(* IEC 61131-3 sources: JingjiangMoonbox/Application/Application/任务列表/Main_Task/IO列表, 15 files *)

(* ---- StEvtReq.st ---- *)
(*@CES
Name=StEvtReq
Type=Gvl
TypeGuid=2db5746d-d284-4425-9f7f-2663a34b0ebc
Guid=8252279d-9d67-4d9b-8f5c-5fb7a358024a
HasDeclaration=True
HasImplementation=False
*)
{DECLARATION}
{attribute 'pack_mode' := '1'}
TYPE StEvtReq :
STRUCT
	xEvt_Estop						: BOOL; (* 急停 *)
	xEvt_Stop						: BOOL; (* 停机 *)
	xEvt_Tension					: BOOL; (* 张力投入 *)
	xEvt_ManuSpdUp					: BOOL; (* 手动加速 *)
	xEvt_ManuSpdDn					: BOOL; (* 手动减速 *)
	xEvt_Ink						: BOOL; (* 空转 *)
	xEvt_Prestart					: BOOL; (* (预)启动 *)
	xEvt_PressAll					: BOOL; (* 全体合压 *)
	xEvt_UnpressAll					: BOOL; (* 全体离压 *)
	xEvt_Print						: BOOL; (* 印刷|联动 *)
	xEvt_AlarmBell					: BOOL; (* 报警 *)
	xEvt_AllInchRun					: BOOL; (* 整机单动 *)
	xEvt_AllExhBlower				: BOOL; (* 整机排风 *)
	xEvt_AllCoolBlower				: BOOL; (* 整机冷风 *)
	xEvt_AllHotBlower				: BOOL; (* 整机热风 *)
	xEvt_AllHeating					: BOOL; (* 整机加热 *)
	xEvt_TapPosition_Printing		: BOOL; (* 2018.7.16.151840/印刷档位 *)
	xEvt_TapPosition_Breaking		: BOOL; (* 2018.7.16.151514/断料档位 *)
	xEvt_TapPosition_UniformInk		: BOOL; (* 2018.7.16.151507/匀墨档位 *)
	xEvt_FastStop					: BOOL;	(* 2022.4.6.110418 快停*)

	xReqEstop						: BOOL; (* 急停 *)
	xReqStop						: BOOL; (* 停机 *)
	xReqTension						: BOOL; (* 张力投入 *)
	xReqManuSpdUp					: BOOL; (* 手动加速 *)
	xReqManuSpdDn					: BOOL; (* 手动减速 *)
	xReqInk							: BOOL; (* 空转 *)
	xReqPrestart					: BOOL; (* (预)启动 *)
	xReqPressAll					: BOOL; (* 全体合压 *)
	xReqUnpressAll					: BOOL; (* 全体离压 *)
	xReqPrint						: BOOL; (* 印刷|联动 *)
	xReqAlarmBell					: BOOL; (* 报警 *)
	xReqAllInchRun					: BOOL; (* 整机单运行 *)
	xReqAllExhBlower				: BOOL; (* 整机排风 *)
	xReqAllCoolBlower				: BOOL; (* 整机冷风 *)
	xReqAllHotBlower				: BOOL; (* 整机热风 *)
	xReqAllHeating					: BOOL; (* 整机加热 *)
	xReqFastStop					: BOOL;	(* 2022.4.6.110418 快停*)
END_STRUCT
END_TYPE

{IMPLEMENTATION}

(* ---- StIOMap_Axis_Extra_FE.st ---- *)
(*@CES
Name=StIOMap_Axis_Extra_FE
Type=Gvl
TypeGuid=2db5746d-d284-4425-9f7f-2663a34b0ebc
Guid=0a3c1562-979e-4c29-a397-fc51d923e0fc
HasDeclaration=True
HasImplementation=False
*)
{DECLARATION}
{attribute 'pack_mode' := '1'}
TYPE StIOMap_Axis_Extra_FE :
STRUCT
	i_xPreHeating							: BOOL; (* 预加热 *)
	i_xPreHeating_Err						: BOOL; (* 预加热报警\温控信号 *)
	i_xPreHotBlower							: BOOL; (* 预热风 *)
	i_xPreHotBlower_Err						: BOOL; (* 预热风报警 *)
	i_xCoolBlower							: BOOL; (* 冷风开关 *)
	i_xCoolBlower_Button					: BOOL; (* 冷风按钮 *)
	i_xCoolBlower_Err						: BOOL; (* 冷风报警 *)
	i_xHotBlower							: BOOL; (* 热风开关 *)
	i_xHotBlower_Button						: BOOL; (* 热风按钮 *)
	i_xHotBlower_Err						: BOOL; (* 热风报警 *)
	i_xHotBlower_Opened_Act					: BOOL; (* 热风实际被打开了|2022.5.11.192858|没有反馈时候需要写true*)
	i_xHotBlower_CHNL2						: BOOL; (* 第2路热风开关 *)
	i_xHotBlower_Button_CHNL2				: BOOL; (* 第2路热风按钮 *)
	i_xHotBlower_Err_CHNL2					: BOOL; (* 第2路热风报警 *)
	i_xHotBlower_Opened_Act_CHNL2			: BOOL; (* 热风2实际被打开了|2022.5.11.192858|没有反馈时候需要写true*)
	i_xTemReachToTarget						: BOOL; (* 到达目标温度 *)
	i_xSteamHeating							: BOOL; (* 蒸汽加热开关 *)
	i_xSteamHeating_Err						: BOOL; (* 蒸汽加热报警 *)
	i_xHeating_I							: BOOL; (* 电加热I档 *)
	i_xHeating_II							: BOOL; (* 电加热II档 *)
	i_xHeating_III							: BOOL; (* 电加热III档 *)
	i_xHeating_Button						: BOOL; (* 加热按钮 *)
	i_xHeating_I_CHNL2						: BOOL; (* 第2路电加热I档 *)
	i_xHeating_II_CHNL2						: BOOL; (* 第2路电加热II档 *)
	i_xHeating_III_CHNL2					: BOOL; (* 第2路电加热III档 *)
	i_xHeating_Button_CHNL2					: BOOL; (* 第2路加热按钮 *)
	i_xAllExhBlower_Up						: BOOL; (* 全上排风 *)
	i_xAllExhBlower_Err_Up					: BOOL; (* 上排风报警 *)
	i_xAllExhBlower_Dn						: BOOL; (* 全下排风 *)
	i_xAllExhBlower_Err_Dn					: BOOL; (* 下排风报警 *)
	i_xAllCoolBlower						: BOOL; (* 全冷风 *)
	i_xAllHotBlower							: BOOL; (* 全热风 *)
	i_xAllHeating							: BOOL; (* 全加热 *)
	i_xAirInletMotorMin_Limit				: BOOL; (* 进风口风门电机最小开度限位 *)
	i_xAirInletMotorMax_Limit				: BOOL; (* 进风口风门电机最大开度限位 *)
	i_xOvensAirOutMotorMin_Limit			: BOOL; (* 烘箱出风口风门电机最小开度限位 *)
	i_xOvensAirOutMotorMax_Limit			: BOOL; (* 烘箱出风口风门电机最大开度限位 *)
	i_xAirExhaustMotorMin_Limit				: BOOL; (* 排风口风门电机最小开度限位 *)
	i_xAirExhaustMotorMax_Limit				: BOOL; (* 排风口风门电机最大开度限位 *)
	i_xAirReturnMotorMin_Limit				: BOOL; (* 回风口风门电机最小开度限位 *)
	i_xAirReturnMotorMax_Limit				: BOOL; (* 回风口风门电机最大开度限位 *)
	i_xScraperInveterError					: BOOL; (* 刮刀变频器报警 *)
	i_xScraperOn							: BOOL; (* 刮刀开关 *)
	i_xInkRollerInveterError				: BOOL; (* 递墨辊变频器报警 |2022.3.26.094940*)
	i_xInkRoller_CW							: BOOL; (* 递墨辊正转开 *)
	i_xInkRoller_CCW						: BOOL; (* 递墨辊反转开 *)
	i_xInkRoller_Up							: BOOL; (* 递墨辊上 *)
	i_xInkRoller_Dn							: BOOL; (* 递墨辊下 *)
	i_xTurnoverFilmAgency					: BOOL; (* 翻料架开关 *)
	i_wAI_AirInletMotor						: WORD; (* 进风口反馈|模拟量控制风门LEL *)
	i_wAI_OvensAirOutMotor					: WORD; (* 烘箱出风口反馈|模拟量控制风门LEL *)
	i_wAI_AirExhaustMotor					: WORD; (* 排风口反馈|模拟量控制风门LEL *)
	i_wAI_AirReturnMotor					: WORD; (* 回风反馈|模拟量控制风门LEL *)
	i_wInputLel								: WORD; (* LEL浓度反馈 *)
	i_wInAllAir								: WORD; (* 总进风反馈输入 *)
	i_wInFreshAir							: WORD; (* 新风反馈输入 *)
	i_wInExhaustAir							: WORD; (* 排风反馈输入 *)
	i_wInReturnAir							: WORD; (* 二次回风反馈输入 *)
	i_xTaper_Incr							: BOOL; (* 增加锥度+|针对牵引 *)
	i_xTaper_Decr							: BOOL; (* 减小锥度-|针对牵引 *)
	i_wAI_CoatingSensor						: WORD; (* 涂布传感器模拟量 *)
	i_byAIType_CoatingSensor				: BYTE; (* 涂布传感器类型 *)
	i_xAirExhaustSwitch						: BOOL; (* 色组排风输入开关 *)
	i_xAirExhaustButton						: BOOL; (* 色组排风输入按钮 *)
	i_xPushIn_PrnRoller						: BOOL; (* 顶版-进 *)
	i_xPullOut_PrnRoller					: BOOL; (* 顶版-退 *)
	i_xRsvd_DI0								: BOOL; (* 数字量输入保留0 *)
	i_xRsvd_DI1								: BOOL; (* 数字量输入保留1 *)
	i_xRsvd_DI2								: BOOL; (* 数字量输入保留2 *)
	i_xRsvd_DI3								: BOOL; (* 数字量输入保留3 *)
	i_xRsvd_DI4								: BOOL; (* 数字量输入保留4 *)
	i_xRsvd_DI5								: BOOL; (* 数字量输入保留5 *)
	i_xRsvd_DI6								: BOOL; (* 数字量输入保留6 *)
	i_xRsvd_DI7								: BOOL; (* 数字量输入保留7 *)
	i_xRsvd_DI8								: BOOL; (* 数字量输入保留8 *)
	i_xRsvd_DI9								: BOOL; (* 数字量输入保留9 *)
	i_xRsvd_DI10							: BOOL; (* 数字量输入保留10 *)
	i_xRsvd_DI11							: BOOL; (* 数字量输入保留11 *)
	i_xRsvd_DI12							: BOOL; (* 数字量输入保留12 *)
	i_xRsvd_DI13							: BOOL; (* 数字量输入保留13 *)
	i_xRsvd_DI14							: BOOL; (* 数字量输入保留14 *)
	i_xRsvd_DI15							: BOOL; (* 数字量输入保留15 *)
	i_wRsvd_AI0								: WORD; (* 模拟量输入保留0 *)
	i_wRsvd_AI1								: WORD; (* 模拟量输入保留1 *)
	i_wRsvd_AI2								: WORD; (* 模拟量输入保留2 *)
	i_wRsvd_AI3								: WORD; (* 模拟量输入保留3 *)
	i_wRsvd_AI4								: WORD; (* 模拟量输入保留4 *)
	i_wRsvd_AI5								: WORD; (* 模拟量输入保留5 *)

	o_xRel_PreHeating						: BOOL; (* 预加热接触器 *)
	o_xLamp_PreHeating						: BOOL; (* 预加热指示灯 *)
	o_xRel_ResetErr_PreHeating				: BOOL; (* 预加热故障复位 *)
	o_wAO_PreHeating						: WORD; (* 预加热模拟量 *)
	o_xRel_PreHeatingRoller_Motor			: BOOL; (* 预热辊使能 *)
	o_xRel_PreHeatingRoller_Motor_Rev		: BOOL; (* 预热辊反转使能 *)
	o_wAO_PreHeatingRoller_Motor			: WORD; (* 预热辊模拟量输出 *)
	o_xRel_PreHotBlower						: BOOL; (* 预热风接触器 *)
	o_xLamp_PreHotBlower					: BOOL; (* 预热风指示灯 *)
	o_xRel_ResetErr_PreHotBlower			: BOOL; (* 预热风故障复位 *)
	o_wAO_PreHotBlower						: WORD; (* 预热风模拟量 *)
	o_xRel_CoolBlower						: BOOL; (* 冷风接触器 *)
	o_xLamp_CoolBlower						: BOOL; (* 冷风指示灯 *)
	o_xRel_HotBlower						: BOOL; (* 热风接触器 *)
	o_xLamp_HotBlower						: BOOL; (* 热风指示灯 *)
	o_xRel_ResetErr_HotBlower				: BOOL; (* 热风故障复位 *)
	o_wAO_HotBlower							: WORD; (* 热风模拟量输出 *)
	o_xRel_HotBlower_CHNL2					: BOOL; (* 第2路热风接触器 *)
	o_xLamp_HotBlower_CHNL2					: BOOL; (* 第2路热风指示灯 *)
	o_xRel_ResetErr_HotBlower_CHNL2			: BOOL; (* 第2路热风故障复位 *)
	o_wAO_HotBlower_CHNL2					: WORD; (* 第2路热风模拟量输出 *)
	o_xRel_SteamHeating						: BOOL; (* 蒸汽输出 *)
	o_xLamp_SteamHeating					: BOOL; (* 蒸汽加热指示灯 *)
	o_xRel_ResetErr_SteamHeating			: BOOL; (* 蒸汽加热复位 *)
	o_wAO_SteamHeating						: WORD; (* 蒸汽加热模拟量输出 *)
	o_xRel_Heating_I						: BOOL; (* 电加热I档 *)
	o_xRel_Heating_II						: BOOL; (* 电加热II档 *)
	o_xRel_Heating_III						: BOOL; (* 电加热III档 *)
	o_xLamp_Heating							: BOOL; (* 电加热指示灯 *)
	o_xRel_Heating_I_CHNL2					: BOOL; (* 第2路电加热I档 *)
	o_xRel_Heating_II_CHNL2					: BOOL; (* 第2路电加热II档 *)
	o_xRel_Heating_III_CHNL2				: BOOL; (* 第2路电加热III档 *)
	o_xLamp_Heating_CHNL2					: BOOL; (* 第2路电加热指示灯 *)
	o_xRel_AllExhBlower_Up					: BOOL; (* 上排风继电器输出 *)
	o_xLamp_AllExhBlower_Up					: BOOL; (* 全上排风指示灯 *)
	o_xRel_ModeStar_AllExhBlower_Up			: BOOL; (* 上排风模式-星形 *)
	o_xRel_ModeTriangle_AllExhBlower_Up		: BOOL; (* 上排风模式-三角 *)
	o_xRel_ResetErr_AllExhBlower_Up			: BOOL; (* 上排风故障复位 *)
	o_wAO_AllExhBlower_Up					: WORD; (* 上排风模拟量输出 *)
	o_xRel_AllExhBlower_Dn					: BOOL; (* 下排风继电器输出 *)
	o_xLamp_AllExhBlower_Dn					: BOOL; (* 全下排风指示灯 *)
	o_xRel_ModeStar_AllExhBlower_Dn			: BOOL; (* 下排风模式-星形 *)
	o_xRel_ModeTriangle_AllExhBlower_Dn		: BOOL; (* 下排风模式-三角 *)
	o_xRel_ResetErr_AllExhBlower_Dn			: BOOL; (* 下排风故障复位 *)
	o_wAO_AllExhBlower_Dn					: WORD; (* 下排风模拟量输出 *)
	o_xLamp_AllCoolBlower					: BOOL; (* 全冷风指示灯 *)
	o_xLamp_AllHotBlower					: BOOL; (* 全热风指示灯 *)
	o_xLamp_AllHeating						: BOOL; (* 全加热指示灯 *)
	o_xAirInletMotor_Increase				: BOOL; (* 进风口风门开度增大 *)
	o_xAirInletMotor_Decrease				: BOOL; (* 进风口风门开度减小 *)
	o_xOvensAirOutMotor_Increase			: BOOL; (* 烘箱出风口风门开度增大 *)
	o_xOvensAirOutMotor_Decrease			: BOOL; (* 烘箱出风口风门开度减小 *)
	o_xAirExhaustMotor_Increase				: BOOL; (* 排风口风门开度增大 *)
	o_xAirExhaustMotor_Decrease				: BOOL; (* 排风口风门开度减小 *)
	o_xAirReturnMotor_Increase				: BOOL; (* 回风风门开度增大 *)
	o_xAirReturnMotor_Decrease				: BOOL; (* 回风风门开度减小 *)
	o_xScraperOn							: BOOL; (* 刮刀输出 *)
(*2022.7.8.093123*)
	o_xScraperRst							: BOOL;(*刮刀故障复位*)
	o_wAO_Scraper							: WORD; (* 刮刀模拟量输出 *)
	o_xInkRollerOn							: BOOL; (* 递墨辊运动信号 *)
	o_xInkRollerRst							: BOOL;(*递墨辊复位2022.7.8.093223*)
	o_xRel_InkRoller_CW						: BOOL; (* 递墨辊正转 *)
	o_xRel_InkRoller_CCW					: BOOL; (* 递墨辊反转 *)
	o_wAO_InkRoller							: WORD; (* 递墨辊模拟量输出 *)
	(*2026.05.25.134825*)
	o_wAO_InkRoller_Dir						:WORD;(*递墨辊模拟量输出@±10V*)
	o_xRel_InkRoller_Up						: BOOL; (* 递墨辊上输出 *)
	o_xRel_InkRoller_Dn						: BOOL; (* 递墨辊下输出 *)
	o_xRel_TurnoverFilmAgency				: BOOL; (* 翻料架输出 *)
	o_xRel_ColdWaterRoller_Motor			: BOOL; (* 水冷辊电机使能 *)
	o_xRel_ColdWaterRoller_Motor_Rev		: BOOL; (* 水冷辊电机反转使能 *)
	o_wAO_ColdWaterRoller_Motor				: WORD; (* 水冷辊电机模拟量输出 *)
	o_xRel_DriveAfterPrint_Motor			: BOOL; (* 印后传动辊电机使能 *)
	o_xRel_DriveAfterPrint_Motor_Rev		: BOOL; (* 印后传动辊电机反转 *)
	o_wAO_DriveAfterPrint_Motor				: WORD; (* 印后传动辊电机模拟量输出 *)
	o_wAO_AirInletMotor						: WORD; (* 进口输出|模拟量控制风门LEL *)
	o_wAO_OvensAirOutMotor					: WORD; (* 烘箱出风口输出|模拟量控制风门LEL *)
	o_wAO_AirExhaustMotor					: WORD; (* 排风口输出|模拟量控制风门LEL *)
	o_wAO_AirReturnMotor					: WORD; (* 回风输出|模拟量控制风门LEL *)
	o_wInAllAir								: WORD; (* 总进风输出 *)
	o_wInFreshAir							: WORD; (* 新风输出 *)
	o_wInExhaustAir							: WORD; (* 排风输出 *)
	o_wInReturnAir							: WORD; (* 二次回风输出 *)
	o_wPreAirHotRollTorque					: WORD; (* 预热辊转矩输出 *)
	o_wCoolWaterRollTorque					: WORD; (* 水冷辊转矩输出 *)
	o_xAirExhaustEn							: BOOL; (* 色组排风输出使能 *)
	o_xRel_PushIn_PrnRoller					: BOOL; (* 顶版-进执行 *)
	o_xRel_PullOut_PrnRoller				: BOOL; (* 顶版-退执行 *)
	o_xRel_ModeStar_HotBlower				: BOOL; (* 热风输出-星形 *)
	o_xRel_ModeTriangle_HotBlower			: BOOL; (* 热风输出-三角 *)
	o_xRel_Oven								: BOOL; (* 色组烘箱输出 *)
	o_xRsvd_DO0								: BOOL; (* 数字量输出保留0 *)
	o_xRsvd_DO1								: BOOL; (* 数字量输出保留1 *)
	o_xRsvd_DO2								: BOOL; (* 数字量输出保留2 *)
	o_xRsvd_DO3								: BOOL; (* 数字量输出保留3 *)
	o_xRsvd_DO4								: BOOL; (* 数字量输出保留4 *)
	o_xRsvd_DO5								: BOOL; (* 数字量输出保留5 *)
	o_xRsvd_DO6								: BOOL; (* 数字量输出保留6 *)
	o_xRsvd_DO7								: BOOL; (* 数字量输出保留7 *)
	o_xRsvd_DO8								: BOOL; (* 数字量输出保留8 *)
	o_xRsvd_DO9								: BOOL; (* 数字量输出保留9 *)
	o_xRsvd_DO10							: BOOL; (* 数字量输出保留10 *)
	o_xRsvd_DO11							: BOOL; (* 数字量输出保留11 *)
	o_xRsvd_DO12							: BOOL; (* 数字量输出保留12 *)
	o_xRsvd_DO13							: BOOL; (* 数字量输出保留13 *)
	o_xRsvd_DO14							: BOOL; (* 数字量输出保留14 *)
	o_xRsvd_DO15							: BOOL; (* 数字量输出保留15 *)
	o_wRsvd_AO0								: WORD; (* 模拟量输出保留0 *)
	o_wRsvd_AO1								: WORD; (* 模拟量输出保留1 *)
	o_wRsvd_AO2								: WORD; (* 模拟量输出保留2 *)
	o_wRsvd_AO3								: WORD; (* 模拟量输出保留3 *)
	o_wRsvd_AO4								: WORD; (* 模拟量输出保留4 *)
	o_wRsvd_AO5								: WORD; (* 模拟量输出保留5 *)
END_STRUCT
END_TYPE

{IMPLEMENTATION}

(* ---- StIOMap_Axis_FE.st ---- *)
(*@CES
Name=StIOMap_Axis_FE
Type=Gvl
TypeGuid=2db5746d-d284-4425-9f7f-2663a34b0ebc
Guid=869f751a-dcb2-42ff-ace2-93e211c33fe9
HasDeclaration=True
HasImplementation=False
*)
{DECLARATION}
{attribute 'pack_mode' := '1'}
TYPE StIOMap_Axis_FE :
STRUCT
	(*IO输入*)
	i_xLinkage								: BOOL; (* 联动 *)
	i_xInch									: BOOL; (* 单运行 *)
	i_xEstop								: BOOL; (* 急停输入 *)
	i_xAlarmBell							: BOOL; (* 警报 *)
	i_xBigAdj								: BOOL; (* 粗调 *)
	i_xLittleAdj							: BOOL; (* 细调 *)
	i_xPressMode_Auto						: BOOL; (* 自动合压 *)
	i_xPressMode_Manu						: BOOL; (* 手动合压 *)
	i_xPress								: BOOL; (* 合压输入 *)
	i_xUnPress								: BOOL; (* 离压输入 *)
	i_xUnPress_Inching						: BOOL; (* 点动离压 *)
	i_xMove_Up								: BOOL; (* 上调 *)
	i_xMove_Down							: BOOL; (* 下调 *)
	i_xMove_Left							: BOOL; (* 左调 *)
	i_xMove_Right							: BOOL; (* 右调 *)
	i_xPosLimit_Left						: BOOL; (* 左限位 *)
	i_xPosLimit_Right						: BOOL; (* 右限位 *)
	i_xHorzMotor_FastSpd					: BOOL; (* 横向电机快 *)
	i_xSleeve_Prn							: BOOL; (* 版辊套筒*)
	i_xSleeve_Net							: BOOL; (* 网辊套筒*)
	i_xPlate_Push_Prn						: BOOL; (* 版辊推出*)
	i_xPlate_Push_Net						: BOOL; (* 网辊推出*)
	i_xAcc									: BOOL; (* 加速 *)
	i_xDec									: BOOL; (* 减速 *)
	i_xInch_Net								: BOOL; (* 网辊单运行-匀墨 *)
		(*2024.09.28.094834//增加秦华IO*)
	i_xJogPaper									: BOOL; (* 走纸点动 *)
	i_xEn_Prn									: BOOL; (* 版辊使能开关 *)

	i_xPrnBigAdj								: BOOL; (* 印刷辊粗调 *)
	i_xPrnLittleAdj								: BOOL; (* 印刷辊细调 *)
	i_xNetBigAdj								: BOOL; (* 网辊粗调 *)
	i_xNetLittleAdj								: BOOL; (* 网辊细调 *)
	i_xStrBigAdj								: BOOL; (* 张带辊粗调 *)
	i_xStrLittleAdj								: BOOL; (* 张带辊细调 *)

	i_xJogUp_Prn_M							: BOOL; (* 印刷辊点动上升 *)
	i_xJogDown_Prn_M						: BOOL; (* 印刷辊点动下降 *)
	i_xJogUp_Prn_G							: BOOL; (* 印刷辊点进上升  传动侧信号*)
	i_xJogDown_Prn_G						: BOOL; (* 印刷辊点动下降  传动侧信号*)
	i_xAllUp_Prn							: BOOL; (* 印刷辊整体上升 *)
	i_xAllDown_Prn							: BOOL; (* 印刷辊整体下降 *)
	i_xJogUp_Str_M							: BOOL; (* 张带辊点动上升 *)
	i_xJogDown_Str_M						: BOOL; (* 张带辊点动下降 *)
	i_xJogUp_Str_G							: BOOL; (* 张带辊点动上升  传动侧信号*)
	i_xJogDown_Str_G						: BOOL; (* 张带辊点动下降  传动侧信号*)
	i_xAllUp_Str							: BOOL; (* 张带辊整体上升 *)
	i_xAllDown_Str							: BOOL; (* 张带辊整体下降 *)
	i_xJogUp_Net_M							: BOOL; (* 网版辊点动前进 *)
	i_xJogDown_Net_M						: BOOL; (* 网版辊点动后退 *)
	i_xJogUp_Net_G							: BOOL; (* 网版辊点动前进 另传动侧信号*)
	i_xJogDown_Net_G						: BOOL; (* 网版辊点动后退  另传动侧信号*)
	i_xAllUp_Net							: BOOL; (* 网版辊整体前进 *)
	i_xAllDown_Net							: BOOL; (* 网版辊整体后退 *)

	i_xSuctionMotor							: BOOL; (* 吸风电机开关*)
	i_xNetMotor								: BOOL;(* 网辊电机开关*)
	i_xNetLock								: BOOL;(* 网辊锁紧开关*)
	i_xStop                             	: BOOL;(* 停止信号*)
	i_xRunning								: BOOL;(* 运行信号*)
	i_xNetPosLimit_Down						: BOOL; (* 网辊下限位 *)
	i_xPrnPosLimit_Up						: BOOL; (* 印刷辊上限位 *)
	i_xPrnPosLimit_Down						: BOOL; (* 印刷辊下限位 *)
	i_xPrnFastUp_M							: BOOL; (* 印刷辊快速上升 *)
	i_xPrnFastDown_M						: BOOL; (* 印刷辊快速下降 *)

	i_xHorzMotor_Alarm						: BOOL;(*横向报警*)
	(*新增变量-开始-wng.nt|2025.08.12.151630*)
	i_xPrnRollerLoose_H						: BOOL;(*夹板报警输入*)
	i_xLostPressure							: BOOL;(*气压低报警*)
	i_xPtcSignal							: BOOL;(*PTC过温报警*)
	(*新增变量-结束-wng.nt|2025.08.12.151630*)

	i_xRsvd_DI0								: BOOL; (* 数字量输入保留0 *)
	i_xRsvd_DI1								: BOOL; (* 数字量输入保留1 *)
	i_xRsvd_DI2								: BOOL; (* 数字量输入保留2 *)
	i_xRsvd_DI3								: BOOL; (* 数字量输入保留3 *)
	i_xRsvd_DI4								: BOOL; (* 数字量输入保留4 *)
	i_xRsvd_DI5								: BOOL; (* 数字量输入保留5 *)
	i_xRsvd_DI6								: BOOL; (* 数字量输入保留6 *)
	i_xRsvd_DI7								: BOOL; (* 数字量输入保留7 *)
	i_xRsvd_DI8								: BOOL; (* 数字量输入保留8 *)
	i_xRsvd_DI9								: BOOL; (* 数字量输入保留9 *)
	i_wRsvd_AI0								: WORD; (* 模拟量输入保留0 *)
	i_wRsvd_AI1								: WORD; (* 模拟量输入保留1 *)
	i_wRsvd_AI2								: WORD; (* 模拟量输入保留2 *)
	i_wRsvd_AI3								: WORD; (* 模拟量输入保留3 *)
	i_wRsvd_AI4								: WORD; (* 模拟量输入保留4 *)
	i_wRsvd_AI5								: WORD; (* 模拟量输入保留5 *)

//IO输出
	o_xLamp_Linkage							: BOOL; (* 色组联动灯 *)
	o_xLamp_Inch							: BOOL; (* 单运行灯 *)
	o_xLamp_Estop							: BOOL; (* 急停灯输出 *)
	o_xLamp_Normal							: BOOL; (* 套色正常 *)
	o_xLamp_Warning							: BOOL; (* 套色报警 *)
	o_xLamp_Lost							: BOOL; (* 套色丢失 *)
	o_xLamp_AxisError						: BOOL; (* 轴故障指示 *)
	o_xRel_ArcAlarm_Unit					: BOOL; (* 本组套色报警输出 *)
	o_xLamp_Press							: BOOL; (* 合压指示 *)
	o_xRel_Press							: BOOL; (* 合压输出 *)
	o_xRel_UnPress							: BOOL; (* 离压输出 *)
	o_xHorzMotor_CW							: BOOL; (* 横向电机正转输出 *)
	o_xHorzMotor_CCW						: BOOL; (* 横向电机反转输出 *)
	o_xRel_Sleeve_Prn						: BOOL; (* 版辊套筒*)
	o_xRel_Sleeve_Net						: BOOL; (* 网辊套筒*)
	o_xRel_Plate_Push_Prn					: BOOL; (* 版辊推出*)
	o_xRel_Plate_Push_Net					: BOOL; (* 网辊推出*)
	o_xLamp_Inch_Net						: BOOL; (* 网辊单动灯 *)
		(*2024.09.28.094834//增加秦华IO*)
	o_xLamp_CorrctionPrn							: BOOL; (* 对版指示灯 *)
	o_xPM_Buzzer_Str								: BOOL; (* 张带辊装版蜂鸣器 *)
	o_xSuctionContactor								: BOOL; (* 吸风接触器 *)
	o_xDamMotorContactor							: BOOL; (* 润板电机接触器 *)
	o_xHydr_station_SV								: BOOL; (* 液压站电磁阀 *)

	(*新增变量-开始-wng.nt|2025.08.12.151630*)
	o_xLamp_Stop							: BOOL;(*停止指示灯*)
	o_xPrnRollerLoose_H						: BOOL;(*夹板报警输入*)
	o_xLostPressure							: BOOL;(*气压低报警*)
	o_xPtcTempHigh							: BOOL;(*PTC过温报警*)
	(*新增变量-结束-wng.nt|2025.08.12.151630*)

	o_xRsvd_DO0								: BOOL; (* 数字量输出保留0 *)
	o_xRsvd_DO1								: BOOL; (* 数字量输出保留1 *)
	o_xRsvd_DO2								: BOOL; (* 数字量输出保留2 *)
	o_xRsvd_DO3								: BOOL; (* 数字量输出保留3 *)
	o_xRsvd_DO4								: BOOL; (* 数字量输出保留4 *)
	o_xRsvd_DO5								: BOOL; (* 数字量输出保留5 *)
	o_xRsvd_DO6								: BOOL; (* 数字量输出保留6 *)
	o_xRsvd_DO7								: BOOL; (* 数字量输出保留7 *)
	o_xRsvd_DO8								: BOOL; (* 数字量输出保留8 *)
	o_xRsvd_DO9								: BOOL; (* 数字量输出保留9 *)
	o_wRsvd_AO0								: WORD; (* 模拟量输出保留0 *)
	o_wRsvd_AO1								: WORD; (* 模拟量输出保留1 *)
	o_wRsvd_AO2								: WORD; (* 模拟量输出保留2 *)
	o_wRsvd_AO3								: WORD; (* 模拟量输出保留3 *)
	o_wRsvd_AO4								: WORD; (* 模拟量输出保留4 *)
	o_wRsvd_AO5								: WORD; (* 模拟量输出保留5 *)
END_STRUCT
END_TYPE

{IMPLEMENTATION}

(* ---- StIOMap_Main_FE.st ---- *)
(*@CES
Name=StIOMap_Main_FE
Type=Gvl
TypeGuid=2db5746d-d284-4425-9f7f-2663a34b0ebc
Guid=2d022e5e-72f6-4cce-877c-3428f23a092c
HasDeclaration=True
HasImplementation=False
*)
{DECLARATION}
{attribute 'pack_mode' := '1'}
TYPE StIOMap_Main_FE :
STRUCT
//(*IO输入*)
	i_xPrestart								: BOOL; //(* 预启动 *)
	i_xInk									: BOOL; //(* 空转 *)
	i_xTension								: BOOL; //(* 张力投入 *)
	i_xPrint								: BOOL; //(* 印刷 *)
	i_xAcc									: BOOL; //(* 加速 *)
	i_xDec									: BOOL; //(* 减速 *)
	i_xPressAll								: BOOL; //(* 全合压 *)
	i_xUnPressAll							: BOOL; //(* 全离压 *)
	i_xEstop								: BOOL; //(* 急停输入 *)
	i_xStop									: BOOL; //(* 停机 *)
	i_xFastStop								: BOOL;(*快停*)
	i_xAlarmBell							: BOOL; //(* 警报 *)
	i_xPressMode_Auto_IF					: BOOL; //(* 放牵自动合压 *)
	i_xPressMode_Manu_IF					: BOOL; //(* 放牵手动合压 *)
	i_xPressMode_Auto_OF					: BOOL; //(* 收牵自动合压 *)
	i_xPressMode_Manu_OF					: BOOL; //(* 收牵手动合压 *)
//2025.12.29.172113增加牵引变频相关变量
	i_xInverterAlarm_If						: BOOL;(*放牵变频报警输入*)
	i_xInverterAlarm_Of						: BOOL;(*收牵变频报警输入*)
	i_xInverterAlarm						: BOOL;(*牵引变频报警输入*)
	i_xInch_If								: BOOL;(*放牵单运行*)
	i_xInch_Of								: BOOL;(*收牵单运行*)

//2023.11.18.135442
	i_xAllExhBlower_Up						: BOOL; (* 全上排风 *)
	i_xAllExhBlower_Err_Up					: BOOL; (* 上排风报警 *)
	i_xAllExhBlower_Dn						: BOOL; (* 全下排风 *)
	i_xAllExhBlower_Err_Dn					: BOOL; (* 下排风报警 *)
	i_xAllCoolBlower						: BOOL; (* 全冷风 *)
	i_xAllHotBlower							: BOOL; (* 全热风 *)
	i_xAllHeating							: BOOL; (* 全加热 *)
	i_xScraperInveterError					: BOOL; (* 刮刀变频器报警 *)
	i_xScraperOn							: BOOL; (* 刮刀开关 *)
	i_xInkRollerInveterError				: BOOL; (* 递墨辊变频器报警 |2022.3.26.094940*)
	i_xInkRoller_CW							: BOOL; (* 递墨辊正转开 *)
	i_xInkRoller_CCW						: BOOL; (* 递墨辊反转开 *)

		(*2024.09.28.094834//增加秦华IO*)
	i_xJumpSelection						: BOOL; (* 跳板选择开关 *)
	i_xHydraulicPower						: BOOL; (* 液压站电源开关 *)
	(*2025.02.25.90543*)
	i_xPressMode_Auto_OF1					: BOOL; //(* 收卷后牵引辊自动合压 *)
	i_xPressMode_Manu_OF1					: BOOL; //(* 收卷后牵引辊手动合压 *)
	i_xTapPosition_Breaking					: BOOL; (* 断料档位 *)
	i_xTapPosition_UniformInk				: BOOL; (* 匀墨档位 *)

	i_xRsvd_DI0								: BOOL; //(* 数字量输入保留0 *)
	i_xRsvd_DI1								: BOOL; //(* 数字量输入保留1 *)
	i_xRsvd_DI2								: BOOL; //(* 数字量输入保留2 *)
	i_xRsvd_DI3								: BOOL; //(* 数字量输入保留3 *)
	i_xRsvd_DI4								: BOOL; //(* 数字量输入保留4 *)
	i_xRsvd_DI5								: BOOL; //(* 数字量输入保留5 *)
	i_xRsvd_DI6								: BOOL; //(* 数字量输入保留6 *)
	i_xRsvd_DI7								: BOOL; //(* 数字量输入保留7 *)
	i_xRsvd_DI8								: BOOL; //(* 数字量输入保留8 *)
	i_xRsvd_DI9								: BOOL; //(* 数字量输入保留9 *)
	i_wRsvd_AI0								: WORD; //(* 模拟量输入保留0 *)
	i_wRsvd_AI1								: WORD; //(* 模拟量输入保留1 *)
	i_wRsvd_AI2								: WORD; //(* 模拟量输入保留2 *)
	i_wRsvd_AI3								: WORD; //(* 模拟量输入保留3 *)
	i_wRsvd_AI4								: WORD; //(* 模拟量输入保留4 *)
	i_wRsvd_AI5								: WORD; //(* 模拟量输入保留5 *)

	o_xLamp_Prestart						: BOOL; //(* 预启动指示 *)
	o_xLamp_Ink								: BOOL; //(* 空转指示 *)
	o_xLamp_Tension							: BOOL; //(* 张力投入指示 *)
	o_xLamp_Print							: BOOL; //(* 印刷指示 *)
	o_xLamp_Acc								: BOOL; //(* 加速指示 *)
	o_xLamp_Dec								: BOOL; //(* 减速指示 *)
	o_xLamp_AllPress						: BOOL; //(* 全合压指示 *)
	o_xLamp_UnPressAll						: BOOL; //(* 全离压指示 *)
	o_xLamp_Estop							: BOOL; //(* 急停灯输出 *)
	o_xLamp_Stop							: BOOL; //(* 指示|停机 *)
	o_xRel_AlarmBell						: BOOL; //(* 报警输出 *)
	o_xRel_ArcAlarm							: BOOL; //(* 整机套色报警输出 *)
	o_xLamp_Press_IF						: BOOL; //(* 放牵合压指示 *)
	o_xRel_Press_IF							: BOOL; //(* 放牵合压输出 *)
	o_xLamp_Press_OF						: BOOL; //(* 收牵合压指示 *)
	o_xRel_Press_OF							: BOOL; //(* 收牵合压输出 *)
//2025.12.29.172304增加	牵引变频控制相关
	o_xCW_If								: BOOL; (* 放牵正转 *)
	o_wAO_If								: WORD; (* 放牵输出频率 *)
	o_xCW_Of								: BOOL; (* 收牵正转 *)
	o_wAO_Of								: WORD; (* 收牵输出频率 *)
	o_xAdjustEn_If							: BOOL; (* 放牵自调使能 *)
	o_wFilm_Vel_If							: WORD; (* 放牵主机速度 *)
	o_xAdjustEn_Of							: BOOL; (* 收牵自调使能 *)
	o_wFilm_Vel_Of							: WORD; (* 收牵主机速度 *)
	o_xINVERTER_RESET						: BOOL; (* (放/收)牵引变频复位 *)
	o_xInverterReset_If						: BOOL; (* 放牵变频复位 *)
	o_xInverterReset_Of						: BOOL; (* 收牵变频复位 *)

//2023.11.18.135519
	o_xRel_AllExhBlower_Up					: BOOL; (* 上排风继电器输出 *)
	o_xLamp_AllExhBlower_Up					: BOOL; (* 全上排风指示灯 *)
	o_xRel_ModeStar_AllExhBlower_Up			: BOOL; (* 上排风模式-星形 *)
	o_xRel_ModeTriangle_AllExhBlower_Up		: BOOL; (* 上排风模式-三角 *)
	o_xRel_ResetErr_AllExhBlower_Up			: BOOL; (* 上排风故障复位 *)
	o_wAO_AllExhBlower_Up					: WORD; (* 上排风模拟量输出 *)
	o_xRel_AllExhBlower_Dn					: BOOL; (* 下排风继电器输出 *)
	o_xLamp_AllExhBlower_Dn					: BOOL; (* 全下排风指示灯 *)
	o_xRel_ModeStar_AllExhBlower_Dn			: BOOL; (* 下排风模式-星形 *)
	o_xRel_ModeTriangle_AllExhBlower_Dn		: BOOL; (* 下排风模式-三角 *)
	o_xRel_ResetErr_AllExhBlower_Dn			: BOOL; (* 下排风故障复位 *)
	o_wAO_AllExhBlower_Dn					: WORD; (* 下排风模拟量输出 *)
	o_xLamp_AllCoolBlower					: BOOL; (* 全冷风指示灯 *)
	o_xLamp_AllHotBlower					: BOOL; (* 全热风指示灯 *)
	o_xLamp_AllHeating						: BOOL; (* 全加热指示灯 *)
 	o_xScraperOn							: BOOL; (* 刮刀输出 *)
(*2022.7.8.093123*)
	o_xScraperRst							: BOOL;(*刮刀故障复位*)
	o_wAO_Scraper							: WORD; (* 刮刀模拟量输出 *)
	o_xInkRollerOn							: BOOL; (* 递墨辊运动信号 *)
	o_xInkRollerRst							: BOOL;(*递墨辊复位2022.7.8.093223*)
	o_xRel_InkRoller_CW						: BOOL; (* 递墨辊正转 *)
	o_xRel_InkRoller_CCW					: BOOL; (* 递墨辊反转 *)
	o_wAO_InkRoller							: WORD; (* 递墨辊模拟量输出 *)

	o_xRsvd_DO0								: BOOL; //(* 数字量输出保留0 *)
	o_xRsvd_DO1								: BOOL; //(* 数字量输出保留1 *)
	o_xRsvd_DO2								: BOOL; //(* 数字量输出保留2 *)
	o_xRsvd_DO3								: BOOL; //(* 数字量输出保留3 *)
	o_xRsvd_DO4								: BOOL; //(* 数字量输出保留4 *)
	o_xRsvd_DO5								: BOOL; //(* 数字量输出保留5 *)
	o_xRsvd_DO6								: BOOL; //(* 数字量输出保留6 *)
	o_xRsvd_DO7								: BOOL; //(* 数字量输出保留7 *)
	o_xRsvd_DO8								: BOOL; //(* 数字量输出保留8 *)
	o_xRsvd_DO9								: BOOL; //(* 数字量输出保留9 *)
	o_wRsvd_AO0								: WORD; //(* 模拟量输出保留0 *)
	o_wRsvd_AO1								: WORD; //(* 模拟量输出保留1 *)
	o_wRsvd_AO2								: WORD; //(* 模拟量输出保留2 *)
	o_wRsvd_AO3								: WORD; //(* 模拟量输出保留3 *)
	o_wRsvd_AO4								: WORD; //(* 模拟量输出保留4 *)
	o_wRsvd_AO5								: WORD; //(* 模拟量输出保留5 *)
END_STRUCT
END_TYPE

{IMPLEMENTATION}

(* ---- StIOMap_UwRw_FE.st ---- *)
(*@CES
Name=StIOMap_UwRw_FE
Type=Gvl
TypeGuid=2db5746d-d284-4425-9f7f-2663a34b0ebc
Guid=f0d92865-0211-4c93-96fb-69cc6a414734
HasDeclaration=True
HasImplementation=False
*)
{DECLARATION}
{attribute 'pack_mode' := '1'}
TYPE StIOMap_UwRw_FE :
STRUCT
	i_xEstop								: BOOL; (* 急停输入 *)
	i_xSafetyGrating						: BOOL; (* 安全光栅 *)
	i_xSafeTyGratingReset					: BOOL;	(* 安全光栅复位*)
	i_xInverterErrorA						: BOOL; (* A轴变频器故障 *)
	i_xInverterErrorB						: BOOL; (* B轴变频器故障 *)
	i_xPreCut								: BOOL; (* 预备接料 *)
	i_xCut_Cancel							: BOOL; (* 接料取消 *)
	i_xCut									: BOOL; (* 接料 *)
	i_xForward								: BOOL; (* 翻转架正转 *)
	i_xReversal								: BOOL; (* 翻转架反转 *)
	i_xAxisExchange							: BOOL; (* 轴切换 *)
(*2021.11.2.161530  替换*)
(**)
(*	i_xCutOnTopKnob							: BOOL; (* 上下裁 |旋钮*)*)
	i_xCutOnTopBtn							: BOOL; (* 上下裁 |按钮*)
	i_xIsUpCut								: BOOL; (* 上裁 *)
	i_xAxisA_Locating_UpCut					: BOOL; (* 上裁A轴定位 *)
	i_xAxisB_Locating_UpCut					: BOOL; (* 上裁B轴定位 *)
	i_xAxisA_Locating_UpCut_PaperCore6Inch	: BOOL; (* 上裁A轴6寸定位 *)
	i_xAxisB_Locating_UpCut_PaperCore6Inch	: BOOL; (* 上裁B轴6寸定位 *)
	i_xMinimumDiamProtect_UpCut				: BOOL; (* 上裁最小卷径保护 *)
	i_xAxisA_MinimumDiamProtect_UpCut		: BOOL; (* 上裁A轴最小卷径保护 *)
	i_xAxisB_MinimumDiamProtect_UpCut		: BOOL; (* 上裁B轴最小卷径保护 *)
	i_xSensor_DiamMeasureLocating_UpCut		: BOOL; (* 上裁卷径测量定位 *)
	i_xSensor_Reflex_UpCut					: BOOL; (* 上裁弧面信号 *)
	i_xAxisA_Locating_DnCut					: BOOL; (* 下裁A轴定位 *)
	i_xAxisB_Locating_DnCut					: BOOL; (* 下裁B轴定位 *)
	i_xAxisA_Locating_DnCut_PaperCore6Inch	: BOOL; (* 下裁A轴6寸定位 *)
	i_xAxisB_Locating_DnCut_PaperCore6Inch	: BOOL; (* 下裁B轴6寸定位 *)
	i_xMinimumDiamProtect_DnCut				: BOOL; (* 下裁最小卷径保护 *)
	i_xAxisB_MinimumDiamProtect_DnCut		: BOOL; (* 下裁A轴最小卷径保护 *)
	i_xAxisA_MinimumDiamProtect_DnCut		: BOOL; (* 下裁B轴最小卷径保护 *)
	i_xSensor_DiamMeasureLocating_DnCut		: BOOL; (* 下裁卷径测量定位 *)
	i_xSensor_Reflex_DnCut					: BOOL; (* 下裁弧面信号 *)
	i_xSensor_Reflex_A_Up						: BOOL; (* A轴弧面信号 *)
	i_xSensor_Reflex_B_Up						: BOOL; (* B轴弧面信号 *)
	i_xSensor_Reflex_A_Dn						: BOOL; (* A轴弧面信号 *)
	i_xSensor_Reflex_B_Dn						: BOOL; (* B轴弧面信号 *)
	i_xPaperCoreSelect6Inch					: BOOL; (* 6寸纸管有效 *)
	i_xInverterManuReset					: BOOL; (* 变频器故障手动复位 *)
	i_xAPos_Mixed							: BOOL; (* 一刀双裁A点位置 *)
	i_xBPos_Mixed							: BOOL; (* 一刀双裁B点位置 *)
	i_xHolderInPosition_Mixed				: BOOL; (* 一刀双裁大臂到位 *)
	i_xTaper_Incr							: BOOL; (* 增加锥度 *)
	i_xTaper_Decr							: BOOL; (* 减小锥度 *)
	i_xAxisInch								: BOOL; (* 轴单运行 |2022.5.24.091430*)
	i_xAxisInch_Rev							: BOOL; (*反向单运行*)
	(*2024.09.28.094834//增加秦华IO*)
	i_xOperation_UWRW						: BOOL; (* 收放卷运行信号 *)
	i_xSynchronous							: BOOL; (* 同步信号 *)
	i_xUwMeasureSensor						: BOOL;(*包含了对射电眼检测和接近开关检测*)
	i_xRsvd_DI0								: BOOL; (* 数字量输入保留0 *)
	i_xRsvd_DI1								: BOOL; (* 数字量输入保留1 *)
	i_xRsvd_DI2								: BOOL; (* 数字量输入保留2 *)
	i_xRsvd_DI3								: BOOL; (* 数字量输入保留3 *)
	i_xRsvd_DI4								: BOOL; (* 数字量输入保留4 *)
	i_xRsvd_DI5								: BOOL; (* 数字量输入保留5 *)
	i_xRsvd_DI6								: BOOL; (* 数字量输入保留6 *)
	i_xRsvd_DI7								: BOOL; (* 数字量输入保留7 *)
	i_xRsvd_DI8								: BOOL; (* 数字量输入保留8 *)
	i_xRsvd_DI9								: BOOL; (* 数字量输入保留9 *)
	i_xRsvd_DI10							: BOOL; (* 数字量输入保留10 *)
	i_xRsvd_DI11							: BOOL; (* 数字量输入保留11 *)
	i_xRsvd_DI12							: BOOL; (* 数字量输入保留12 *)
	i_xRsvd_DI13							: BOOL; (* 数字量输入保留13 *)
	i_xRsvd_DI14							: BOOL; (* 数字量输入保留14 *)
	i_xRsvd_DI15							: BOOL; (* 数字量输入保留15 *)
	i_wRsvd_AI0								: WORD; (* 模拟量输入保留0 *)
	i_wRsvd_AI1								: WORD; (* 模拟量输入保留1 *)
	i_wRsvd_AI2								: WORD; (* 模拟量输入保留2 *)
	i_wRsvd_AI3								: WORD; (* 模拟量输入保留3 *)
	i_wRsvd_AI4								: WORD; (* 模拟量输入保留4 *)
	i_wRsvd_AI5								: WORD; (* 模拟量输入保留5 *)

	o_xEstopLamp							: BOOL; (* 急停指示 *)
	o_xLamp_SafeTyGrating					: BOOL;	(* 安全光栅触发灯|有光栅输入时候输出*)
	o_xRel_AlarmBell						: BOOL; (* 警铃输出 *)
	o_xInverterResetA						: BOOL; (* A轴变频复位 *)
	o_xInverterResetB						: BOOL; (* B轴变频复位 *)
	o_xLamp_InverterError_A					: BOOL; (* A轴变频故障指示 *)
	o_xLamp_InverterError_B					: BOOL; (* B轴变频故障指示 *)
	o_xInverterReset_ALL					: BOOL; (* 变频器整体复位 *)
	o_xLamp_InverterError_ALL				: BOOL; (* 整机变频故障指示 *)
	o_xLamp_PreDrive						: BOOL; (* 预驱同步指示 *)
	o_xRel_TowerForeward					: BOOL; (* 塔台正转 *)
	o_xRel_TowerReversal					: BOOL; (* 塔台反转 *)
	o_xAxisALamp							: BOOL; (* A轴指示 *)
	o_xAxisBLamp							: BOOL; (* B轴指示 *)
	o_xAxisAForeward						: BOOL; (* A轴正转 *)
	o_xAxisAReversal						: BOOL; (* A轴反转 *)
	o_xAxisAZeroServo						: BOOL; (* A轴零伺服 *)
	o_xAxisBForeward						: BOOL; (* B轴正转 *)
	o_xAxisBReversal						: BOOL; (* B轴反转 *)
	o_xAxisBZeroServo						: BOOL; (* B轴零伺服 *)
	o_xCutOnTop								: BOOL; (* 上裁刀-反之代表下裁刀*)
	o_xCutHolder_UpCut						: BOOL; (* 上裁刀架 *)
	o_xCutCylinder_UpCut					: BOOL; (* 上裁胶辊 *)
	o_xCutter_UpCut							: BOOL; (* 上裁裁刀 *)
	o_xCutHolder_DnCut						: BOOL; (* 下裁刀架 *)
	o_xCutCylinder_DnCut					: BOOL; (* 下裁胶辊 *)
	o_xCutter_DnCut							: BOOL; (* 下裁裁刀 *)
	o_xLamp_PaperCoreSelect6Inch			: BOOL; (* 6寸纸管指示 *)
	o_xLamp_InverterError					: BOOL; (* 变频器故障指示 *)
	o_xRel_HolderCylinder_Up_Mixed			: BOOL; (* 一刀双裁大臂气缸-上 *)
	o_xRel_RollerCylinder_Up_Mixed			: BOOL; (* 一刀双裁胶辊气缸-上 *)
	o_xRel_CutterCylinder_Up_Mixed			: BOOL; (* 一刀双裁裁刀气缸-上 *)
	o_xRel_HolderCylinder_Dn_Mixed			: BOOL; (* 一刀双裁大臂气缸-下 *)
	o_xRel_RollerCylinder_Dn_Mixed			: BOOL; (* 一刀双裁胶辊气缸-下 *)
	o_xRel_CutterCylinder_Dn_Mixed			: BOOL; (* 一刀双裁裁刀气缸-下 *)
	o_xRel_TowerForeward_Mixed				: BOOL; (* 一刀双裁塔台正转 *)
	o_xRel_TowerReversal_Mixed				: BOOL; (* 一刀双裁塔台反转 *)
	o_xAxisATorqueCancel					: BOOL; (* A轴转矩取消 *)
	o_xAxisBTorqueCancel					: BOOL; (* B轴转矩取消 *)
	o_wAxisATorqueVolt						: WORD; (* A轴转矩电压 *)
	o_wAxisBTorqueVolt						: WORD; (* B轴转矩电压 *)
	o_xLampAxisInching						: BOOL; (* 轴单运行中*)
	(*2024.09.28.094834//增加秦华IO*)
	o_xHydrPumpPower						: BOOL; (* 液压泵电源开关 *)
	o_xAdvanceAllBoot						: BOOL; (* 开机整体进版信号 *)
	o_xStopBack								: BOOL; (* 停止退版信号 *)
	o_xOutputAlarm							: BOOL; (* 警报输出 *)
	o_xLampInk								: BOOL; (* 空转信号 *)
	o_xServoError							: BOOL; (* 伺服故障信号 *)
	o_xRsvd_DO0								: BOOL; (* 数字量输出保留0 *)
	o_xRsvd_DO1								: BOOL; (* 数字量输出保留1 *)
	o_xRsvd_DO2								: BOOL; (* 数字量输出保留2 *)
	o_xRsvd_DO3								: BOOL; (* 数字量输出保留3 *)
	o_xRsvd_DO4								: BOOL; (* 数字量输出保留4 *)
	o_xRsvd_DO5								: BOOL; (* 数字量输出保留5 *)
	o_xRsvd_DO6								: BOOL; (* 数字量输出保留6 *)
	o_xRsvd_DO7								: BOOL; (* 数字量输出保留7 *)
	o_xRsvd_DO8								: BOOL; (* 数字量输出保留8 *)
	o_xRsvd_DO9								: BOOL; (* 数字量输出保留9 *)
	o_xRsvd_DO10							: BOOL; (* 数字量输出保留10 *)
	o_xRsvd_DO11							: BOOL; (* 数字量输出保留11 *)
	o_xRsvd_DO12							: BOOL; (* 数字量输出保留12 *)
	o_xRsvd_DO13							: BOOL; (* 数字量输出保留13 *)
	o_xRsvd_DO14							: BOOL; (* 数字量输出保留14 *)
	o_xRsvd_DO15							: BOOL; (* 数字量输出保留15 *)
	o_wRsvd_AO0								: WORD; (* 模拟量输出保留0 *)
	o_wRsvd_AO1								: WORD; (* 模拟量输出保留1 *)
	o_wRsvd_AO2								: WORD; (* 模拟量输出保留2 *)
	o_wRsvd_AO3								: WORD; (* 模拟量输出保留3 *)
	o_wRsvd_AO4								: WORD; (* 模拟量输出保留4 *)
	o_wRsvd_AO5								: WORD; (* 模拟量输出保留5 *)
END_STRUCT
END_TYPE

{IMPLEMENTATION}

(* ---- StProgMonitoring.st ---- *)
(*@CES
Name=StProgMonitoring
Type=Gvl
TypeGuid=2db5746d-d284-4425-9f7f-2663a34b0ebc
Guid=212a47fe-cf90-4c52-849d-68b6b927c1da
HasDeclaration=True
HasImplementation=False
*)
{DECLARATION}
{attribute 'pack_mode' := '1'}
TYPE StProgMonitoring :
STRUCT
	i_lrUw_real				: LREAL; (* 放料摆臂真实值/2019.1.25.091316 *)
	i_lrUw_cur				: LREAL; (* 放料摆臂电压值/相对中位 *)
	i_wUw_cur				: WORD; (* 放料摆臂数字值 *)
	i_lrIf_real				: LREAL; (* 放牵摆臂真实值/2019.1.25.091307 *)
	i_lrIf_cur				: LREAL; (* 放牵摆臂电压值/相对中位 *)
	i_wIf_cur				: WORD; (* 放牵摆臂数字值 *)
	i_lrOf_real				: LREAL; (* 收牵摆臂真实值/2019.1.25.091256 *)
	i_lrOf_cur				: LREAL; (* 收牵摆臂电压值/相对中位 *)
	i_wOf_cur				: WORD; (* 收牵摆臂数字值 *)
	i_lrRw_real				: LREAL; (* 收料摆臂真实值/2019.1.25.091233 *)
	i_lrRw_cur				: LREAL; (* 收料摆臂数字值/相对中位 *)
	i_wRw_cur				: WORD; (* 收料摆臂电压值 *)
	i_lrPressure_Vol		: LREAL; (* 压力传感器电压值 *)
	i_wPressure_Vol			: WORD; (* 压力传感器数字值 *)
	o_wUwAxisA_cur			: WORD; (* 放料A轴数值 *)
	o_lrUwAxisA_Vol			: LREAL; (* 放料A轴电压值 *)
	o_lrUwAxisA_Feq			: LREAL; (* 放料A轴频率 *)
	o_wUwAxisB_cur			: WORD; (* 放料B轴数值 *)
	o_lrUwAxisB_Vol			: LREAL; (* 放料B轴电压值 *)
	o_lrUwAxisB_Feq			: LREAL; (* 放料B轴频率 *)
	o_wRwAxisA_cur			: WORD; (* 收料A轴数值 *)
	o_lrRwAxisA_Vol			: LREAL; (* 收料A轴电压值 *)
	o_lrRwAxisA_Feq			: LREAL; (* 收料A轴频率 *)
	o_wRwAxisB_cur			: WORD; (* 收料B轴数值 *)
	o_lrRwAxisB_Vol			: LREAL; (* 收料B轴电压值 *)
	o_lrRwAxisB_Feq			: LREAL; (* 收料B轴频率 *)
	o_wVelocity_cur			: WORD; (* 线速度表数值 *)
	o_lrVelocity_Vol		: LREAL; (* 线速度表电压值 *)
	o_wTaper_cur			: WORD; (* 电控比例阀数值 *)
	o_lrTaper_Vol			: LREAL; (* 电控比例阀电压值 *)
	o_wIf_cur				: WORD; (* 放牵数值 *)
	o_lrIf_Vol				: LREAL; (* 放牵电压值 *)
	o_lrIf_Feq				: LREAL; (* 放牵频率 *)
	o_wOf_cur				: WORD; (* 收牵数值 *)
	o_lrOf_Vol				: LREAL; (* 收牵电压值 *)
	o_lrOf_Feq				: LREAL; (* 收牵频率 *)
	o_wPreHotRoller_Vol		: WORD; (* 传动辊/预热辊数字值 *)
	o_lrPreHotRoller_Vol	: LREAL; (* 传动辊/预热辊电压值 *)
	i_wDiamMeasureUpCut		: WORD; (* 上裁卷径电位器/2018.11.22.103723 *)
	i_lrDiamMeasureUpCut	: LREAL; (* 上裁卷径电位器/2018.11.22.103723 *)
	i_wDiamMeasureDnCut		: WORD; (* 下裁卷径电位器/2018.11.22.103730 *)
	i_lrDiamMeasureDnCut	: LREAL; (* 上裁卷径电位器/2018.11.22.103723 *)

	(*2023.09.04.144717@20bytes*)
	i_wDiamMeasureAxisA		: WORD; (* A轴卷径超声波/ *)
	i_lrDiamMeasureAxisA	: LREAL; (* A轴卷径超声波/*)
	i_wDiamMeasureAxisB		: WORD; (* B轴卷径超声波/*)
	i_lrDiamMeasureAxisB	: LREAL; (* B轴卷径超声波/*)
	abyReservedFields		: ARRAY [1..20] OF BYTE; (* 预留空间 *)
END_STRUCT
END_TYPE

{IMPLEMENTATION}

(* ---- KS_InitStEvtReq.st ---- *)
(*@CES
Name=KS_InitStEvtReq
Type=FunctionBlock
TypeGuid=6f9dac99-8de1-4efc-8465-68ac443b7d08
Guid=29056b31-c015-4828-ae2e-3b4c94234de1
HasDeclaration=True
HasImplementation=True
*)
{DECLARATION}
FUNCTION KS_InitStEvtReq : INT
VAR_INPUT
	i_pstStEvtReq: POINTER TO StEvtReq;
END_VAR
VAR
	iResult: INT;
END_VAR
{IMPLEMENTATION}
iResult:= 0;
IF i_pstStEvtReq<>0 THEN
	i_pstStEvtReq^.xEvt_Estop:= FALSE; (* 急停 *)
	i_pstStEvtReq^.xEvt_Stop:= FALSE; (* 停机 *)
	i_pstStEvtReq^.xEvt_FastStop:= FALSE; (* 快速停机 *)
	i_pstStEvtReq^.xEvt_Tension:= FALSE; (* 张力投入 *)
	i_pstStEvtReq^.xEvt_ManuSpdUp:= FALSE; (* 手动加速 *)
	i_pstStEvtReq^.xEvt_ManuSpdDn:= FALSE; (* 手动减速 *)
	i_pstStEvtReq^.xEvt_Ink:= FALSE; (* 空转 *)
	i_pstStEvtReq^.xEvt_Prestart:= FALSE; (* (预)启动 *)
	i_pstStEvtReq^.xEvt_PressAll:= FALSE; (* 全体合压 *)
	i_pstStEvtReq^.xEvt_UnpressAll:= FALSE; (* 全体离压 *)
	i_pstStEvtReq^.xEvt_Print:= FALSE; (* 印刷/联动 *)
	i_pstStEvtReq^.xEvt_AlarmBell:= FALSE; (* 报警 *)
	i_pstStEvtReq^.xEvt_AllInchRun:= FALSE; (* 整机单动 *)
	i_pstStEvtReq^.xEvt_AllExhBlower:= FALSE; (* 排风启动 *)
	i_pstStEvtReq^.xEvt_AllCoolBlower:= FALSE; (* 2018.7.19.142033/冷风启动 *)
	i_pstStEvtReq^.xEvt_AllHotBlower:= FALSE; (* 热风启动 *)
	i_pstStEvtReq^.xEvt_AllHeating:= FALSE; (* 加热启动 *)
	i_pstStEvtReq^.xEvt_TapPosition_Printing:= FALSE; (* 2018.7.16.151840/印刷档位 *)
	i_pstStEvtReq^.xEvt_TapPosition_Breaking:= FALSE; (* 2018.7.16.151514/断料档位 *)
	i_pstStEvtReq^.xEvt_TapPosition_UniformInk:= FALSE; (* 2018.7.16.151507/匀墨档位 *)

	i_pstStEvtReq^.xReqEstop:= FALSE; (* 急停 *)
	i_pstStEvtReq^.xReqStop:= FALSE; (* 停机 *)
	i_pstStEvtReq^.xReqFastStop:= FALSE; (* 快速停机 *)
	i_pstStEvtReq^.xReqTension:= FALSE; (* 张力投入 *)
	i_pstStEvtReq^.xReqManuSpdUp:= FALSE; (* 手动加速 *)
	i_pstStEvtReq^.xReqManuSpdDn:= FALSE; (* 手动减速 *)
	i_pstStEvtReq^.xReqInk:= FALSE; (* 空转 *)
	i_pstStEvtReq^.xReqPrestart:= FALSE; (* (预)启动 *)
	i_pstStEvtReq^.xReqPressAll:= FALSE; (* 全体合压 *)
	i_pstStEvtReq^.xReqUnpressAll:= FALSE; (* 全体离压 *)
	i_pstStEvtReq^.xReqPrint:= FALSE; (* 印刷/联动 *)
	i_pstStEvtReq^.xReqAlarmBell:= FALSE; (* 报警 *)
	i_pstStEvtReq^.xReqAllInchRun:= FALSE; (* 整机单动 *)
	i_pstStEvtReq^.xReqAllExhBlower:= FALSE; (* 整机排风 *)
	i_pstStEvtReq^.xReqAllCoolBlower:= FALSE; (* 整机冷风 *)
	i_pstStEvtReq^.xReqAllHotBlower:= FALSE; (* 整机热风 *)
	i_pstStEvtReq^.xReqAllHeating:= FALSE; (* 整机加热 *)
ELSE
	iResult:= -1;
END_IF

KS_InitStEvtReq:= iResult;

(* ---- KS_QueryRangeByAType.st ---- *)
(*@CES
Name=KS_QueryRangeByAType
Type=FunctionBlock
TypeGuid=6f9dac99-8de1-4efc-8465-68ac443b7d08
Guid=eff421d0-eb21-45f6-be1b-43a1b515e8bd
HasDeclaration=True
HasImplementation=True
*)
{DECLARATION}
FUNCTION KS_QueryRangeByAType : INT
VAR_INPUT
	i_byType_AnglogIO: BYTE; (* 1:0~10v; 2:4~20mA; 3:-5~5v; 4:0~5v; 5:0~20mA/ 0:-10v~10v(默认)*)
	i_plrRange_Min: POINTER TO LREAL;
	i_plrRange_Max: POINTER TO LREAL;
	i_pdiRange_Min: POINTER TO DINT;
	i_pdiRange_Max: POINTER TO DINT;
END_VAR
VAR
	lrN_min: LREAL;
	lrN_max: LREAL;
	diN_min: DINT;
	diN_max: DINT;
END_VAR
{IMPLEMENTATION}
CASE i_byType_AnglogIO OF
1:(*0~10v|*)
	lrN_min:= 0;
	lrN_max:= 10;
	diN_min:= 0;
	diN_max:= 32767;
2:(*4~20mA|*)
	lrN_min:= 4;
	lrN_max:= 20;
	diN_min:= 6553(*0*); (* 修复xie.gc测试lel时期更新的问题|@2020.12.19.101658 *)
	diN_max:= 32767;

3:(*-5~5v|*)
	lrN_min:= -5;
	lrN_max:= 5;
	diN_min:= -32767;
	diN_max:= 32767;
4:(*0~5v|*)
	lrN_min:= 0;
	lrN_max:= 5;
	diN_min:= 0;
	diN_max:= 32767;
5:(*0~20mA|*)
	lrN_min:= 0;
	lrN_max:= 20;
	diN_min:= 0;
	diN_max:= 32767;
ELSE(*所有默认就当正负10v处理|*)
	lrN_min:= -10;
	lrN_max:= 10;
	diN_min:= -32767;
	diN_max:= 32767;
END_CASE

IF i_plrRange_Min<>0 THEN
	i_plrRange_Min^:= lrN_min;
END_IF
IF i_plrRange_Max<>0 THEN
	i_plrRange_Max^:= lrN_max;
END_IF
IF i_pdiRange_Min<>0 THEN
	i_pdiRange_Min^:= diN_min;
END_IF
IF i_pdiRange_Max<>0 THEN
	i_pdiRange_Max^:= diN_max;
END_IF

KS_QueryRangeByAType:= 0;

(* ---- KS_SetValueByAIType.st ---- *)
(*@CES
Name=KS_SetValueByAIType
Type=FunctionBlock
TypeGuid=6f9dac99-8de1-4efc-8465-68ac443b7d08
Guid=1789f748-e9c1-482e-88f3-0e0eb31b2a1c
HasDeclaration=True
HasImplementation=True
*)
{DECLARATION}
FUNCTION KS_SetValueByAIType : BOOL(*根据传感器类型写入换算值|电位器写入模拟量值|绝对值编码器方式根据标志写入绝对值或者换算值*)
(*针对编码器过圈问题处理*)
(*2024.01.21.105453 过圈的处理不太完善*)
VAR_INPUT
	i_dwAIData:DWORD;(*采样值*)
	i_byAiType:BYTE;
	(* 控制0~5的状态切换/0:-10v~10v; /.1:0~10v; /.2:4~20mA; /.3:-5~5v; /.4:0~5v; /.5:0~20mA *)
	(*2022.8.29.174810 增加一种类型|/.6 绝对值编码器方式*)
	i_byOutType:BYTE;(*绝对值方式下输出形式|0: 实际绝对值|1:根据+-10v转换值-相对于中位值的(用于最终计算张力调整量)
					   电位器方式下输出形式|0: 实际值|1:相对于中位值的(用于最终计算张力调整量)*)
	i_lrAIData_med:LREAL;(*中位值*)
	(*2024.01.21.102636 该值应该是编码器旋转的最大角度@以前的注释有问题*)
	i_byMaxAngle_AITypeEnc:BYTE:=60;(*绝对值方式下摆臂最大角度(对称|单位°)|用于控制i_byOutType=1时+-10v和角度对应关系*)
	i_dwEncResolution:DWORD:=8388608;(*单圈分辨率|23BITS*)
	i_plrValue:POINTER TO LREAL;(*换算值*)
END_VAR
VAR
	lrAngle_Med									: LREAL;(*中位角度|0对应0°|i_dwEncResolution对应360°*)
	lrAngle_Cur									: LREAL;(*当前角度|0对应0°|i_dwEncResolution对应360°*)
	lrAngle_Max									: LREAL;(*最大角度(正角度)|相对于中位*)
	lrAngle_Min									: LREAL;(*最小角度(负角度)|相对于中位*)
	iAngle_Max_Valid							: INT:=180;(*最大合法偏摆角度*)
	iAngle_add									: INT:=20;(*在最大角度和最小角度上叠加的角度@这个之内都是合法的*)
	lrN_min										: LREAL;
	lrN_max										: LREAL;
	diN_min										: DINT;
	diN_max										: DINT;
	lrTempResult								: LREAL;
	lrTemp										: LREAL;
	lrTemp1										: LREAL;
	wAIData										: WORD;
END_VAR
{IMPLEMENTATION}
CASE i_byAiType OF
 		6:(*绝对值方式*)
			(*0对应0°|i_dwEncResolution对应360°*)
			IF i_dwEncResolution<>0 THEN
				lrAngle_Cur:=DWORD_TO_LREAL(i_dwAIData)/i_dwEncResolution*360;
			END_IF
			(*0对应0°|i_dwEncResolution对应360°*)
			IF i_dwEncResolution<>0 THEN
				lrAngle_Med:=(i_lrAIData_med)/i_dwEncResolution*360;
			END_IF
			(*求最大\小偏摆角度*)
			lrTemp:=BYTE_TO_LREAL(i_byMaxAngle_AITypeEnc)/2;(*取输入最大摆动的一半|该值在下面运算被使用了*)
			(*计算合法角度范围@2024.01.21.103626+注释*)
			lrAngle_Max:=lrTemp+lrAngle_Med;
			lrAngle_Max:=lrAngle_Max+iAngle_add;(*叠加冗余@2024.01.21.103531*)

			lrAngle_Min:=-lrTemp+lrAngle_Med;
			lrAngle_Min:=lrAngle_Min-iAngle_add;(*叠加冗余@2024.01.21.103528*)

			IF i_byOutType=1 THEN(*转换为+-10V(相对于中位)|-10 对应lrAngle_Min角度|10对应lrAngle_Max角度*)
				IF (lrAngle_Cur>=lrAngle_Min AND
					lrAngle_Cur<=lrAngle_Max) THEN(*当前角度处于区间内*)
					lrTemp1:=lrAngle_Cur-lrAngle_Med;(*相对于中位*)
				ELSIF lrAngle_Cur<lrAngle_Min THEN
					lrTemp1:=lrAngle_Cur+360-lrAngle_Med;(*相对于中位*)
				ELSIF lrAngle_Cur>=lrAngle_Max THEN
					lrTemp1:=lrAngle_Cur-360-lrAngle_Med;(*相对于中位*)
				END_IF

				IF lrTemp<>0 THEN
					lrTempResult:=10/lrTemp*lrTemp1;(*相对于中位值*)
					IF lrTempResult>10 THEN
						lrTempResult:=10;
					ELSIF lrTempResult<=-10 THEN
						lrTempResult:=-10;
					END_IF
				END_IF

			ELSE(*使用当前值*)
				lrTempResult:=DWORD_TO_LREAL(i_dwAIData);
			END_IF

ELSE(*电位器方式*)
	wAIData:=DWORD_TO_WORD(i_dwAIData);
	KS_QueryRangeByAType(i_byAiType, ADR(lrN_min), ADR(lrN_max), ADR(diN_min), ADR(diN_max));
	lrTempResult:= KSIO_DA(WORD_TO_INT(wAIData), lrN_min, lrN_max, diN_min, diN_max);

	IF i_byOutType=1 THEN(*相对于中位值的(用于最终计算张力调整量)*)
		lrTempResult:=lrTempResult-i_lrAIData_med;
	ELSE(*实际值*);
	END_IF
END_CASE

IF i_plrValue<>0 THEN
	i_plrValue^:=lrTempResult;
END_IF

(* ---- KSIO_AD.st ---- *)
(*@CES
Name=KSIO_AD
Type=FunctionBlock
TypeGuid=6f9dac99-8de1-4efc-8465-68ac443b7d08
Guid=aa598b09-6eb3-4e37-bb94-f4d8224e5ed0
HasDeclaration=True
HasImplementation=True
*)
{DECLARATION}
FUNCTION KSIO_AD : DINT
VAR_INPUT
	i_lrVolt: LREAL; (* 电压值 *)
	i_lrVolt_min: LREAL; (* 模拟量量程下限 *)
	i_lrVolt_max: LREAL; (* 模拟量量程上限 *)
	i_diRange_min: DINT; (* 数字量量程下限 *)
	i_diRange_max: DINT; (* 数字量量程上限 *)
END_VAR
VAR
	diResult: DINT;
	diRange_min: DINT;
	diRange_max: DINT;
END_VAR
{IMPLEMENTATION}
diResult:= 0;
IF i_lrVolt_min<>i_lrVolt_max THEN (*分母不能为0*)
	diResult:= LREAL_TO_DINT(i_diRange_min+(i_lrVolt-i_lrVolt_min)*(i_diRange_max-i_diRange_min)/(i_lrVolt_max-i_lrVolt_min)); (*计算实际的数字量*)

	(*取边界值*)
	IF i_diRange_max>=i_diRange_min THEN
		diRange_max:= i_diRange_max;
		diRange_min:= i_diRange_min;
	ELSE
		diRange_max:= i_diRange_min;
		diRange_min:= i_diRange_max;
	END_IF

	(*防止越界||*)
	IF diResult>diRange_max THEN
		diResult:= diRange_max;
	ELSIF diResult<diRange_min THEN
		diResult:= diRange_min;
	END_IF
END_IF

KSIO_AD:= diResult;

(* ---- KSIO_DA.st ---- *)
(*@CES
Name=KSIO_DA
Type=FunctionBlock
TypeGuid=6f9dac99-8de1-4efc-8465-68ac443b7d08
Guid=6e901fa2-602f-4438-9b06-80acf888523a
HasDeclaration=True
HasImplementation=True
*)
{DECLARATION}
FUNCTION KSIO_DA : LREAL
VAR_INPUT
	i_iData: INT; (* 数值输入/由于发现外部使用时直接WORD_TO_DINT()造成边界错误/修复输入类型/2020.1.2.093534_ *)
	i_lrVolt_min: LREAL; (* 模拟量量程下限 *)
	i_lrVolt_max: LREAL; (* 模拟量量程上限 *)
	i_diRange_min: DINT; (* 数字量量程下限 *)
	i_diRange_max: DINT; (* 数字量量程上限 *)
END_VAR
VAR
	lrVolt_min: LREAL;
	lrVolt_max: LREAL;
	lrResult: LREAL;
	diTmpData: DINT; (* 2020.1.2.093627_ *)
END_VAR
{IMPLEMENTATION}
lrResult:= 0;
diTmpData:= INT_TO_DINT(i_iData); (* 2020.1.2.093707_ *)
IF i_diRange_min<>i_diRange_max THEN (* 分母不能为0 *)
	lrResult:= i_lrVolt_min+(diTmpData-i_diRange_min)*(i_lrVolt_max-i_lrVolt_min)/(i_diRange_max-i_diRange_min); (* 计算实际的电压值 *)

	(* 取边界值 *)
	IF i_lrVolt_max>=i_lrVolt_min THEN
		lrVolt_max:= i_lrVolt_max;
		lrVolt_min:= i_lrVolt_min;
	ELSE
		lrVolt_max:= i_lrVolt_min;
		lrVolt_min:= i_lrVolt_max;
	END_IF

	(* 如果超边界就取边界值好了 *)
	IF lrResult>lrVolt_max THEN
		lrResult:= lrVolt_max;
	ELSIF lrResult<lrVolt_min THEN
		lrResult:= lrVolt_min;
	END_IF
END_IF

KSIO_DA:= lrResult;

(* ---- KS_FB_MapAxisIOBasic.st ---- *)
(*@CES
Name=KS_FB_MapAxisIOBasic
Type=FunctionBlock
TypeGuid=6f9dac99-8de1-4efc-8465-68ac443b7d08
Guid=d9b432ef-d857-456a-9063-33429bf446aa
HasDeclaration=True
HasImplementation=True
*)
{DECLARATION}
FUNCTION_BLOCK KS_FB_MapAxisIOBasic
VAR_INPUT
	i_xEn									: BOOL;(*功能块使能|*)
	i_xEnableInput							: BOOL;(*使能输入|*)
	i_xEnableOutput							: BOOL;(*使能输出|*)
	i_pstStIOMap_Axis_FE					: POINTER TO StIOMap_Axis_FE;(*轴io数据区域|*)
	i_xLinkage								: BOOL; (* 联动 *)
	i_xInch									: BOOL; (* 单运行 *)
	i_xEstop								: BOOL; (* 急停输入 *)
	i_xAlarmBell							: BOOL; (* 警报 *)
	i_xBigAdj								: BOOL; (* 粗调 *)
	i_xLittleAdj							: BOOL; (* 细调 *)
	i_xPressMode_Auto						: BOOL; (* 自动合压 *)
	i_xPressMode_Manu						: BOOL; (* 手动合压 *)
	i_xPress								: BOOL; (* 合压输入 *)
	i_xUnPress								: BOOL; (* 离压输入 *)
	i_xUnPress_Inching						: BOOL; (* 点动离压 *)
	i_xMove_Up								: BOOL; (* 上调 *)
	i_xMove_Down							: BOOL; (* 下调 *)
	i_xMove_Left							: BOOL; (* 左调 *)
	i_xMove_Right							: BOOL; (* 右调 *)
	i_xPosLimit_Left						: BOOL; (* 左限位 *)
	i_xPosLimit_Right						: BOOL; (* 右限位 *)
	i_xHorzMotor_FastSpd					: BOOL; (* 横向电机快 *)
	i_xSleeve_Prn							: BOOL; (* 版辊套筒*)
	i_xSleeve_Net							: BOOL; (* 网辊套筒*)
	i_xPlate_Push_Prn						: BOOL; (* 版辊推出*)
	i_xPlate_Push_Net						: BOOL; (* 网辊推出*)
	i_xAcc									: BOOL; (* 加速 *)
	i_xDec									: BOOL; (* 减速 *)
	i_xInch_Net								: BOOL; (* 网辊单运行-匀墨 *)

	(*2024.09.28.094834//增加秦华IO*)
	i_xJogPaper									: BOOL; (* 走纸点动 *)
	i_xEn_Prn									: BOOL; (* 版辊使能开关 *)

	i_xPrnBigAdj								: BOOL; (* 印刷辊粗调 *)
	i_xPrnLittleAdj								: BOOL; (* 印刷辊细调 *)
	i_xNetBigAdj									: BOOL; (* 网辊粗调 *)
	i_xNetLittleAdj								: BOOL; (* 网辊细调 *)
	i_xStrBigAdj								: BOOL; (* 张带辊粗调 *)
	i_xStrLittleAdj								: BOOL; (* 张带辊细调 *)

	i_xJogUp_Prn_M							: BOOL; (* 印刷辊点动上升 *)
	i_xJogDown_Prn_M						: BOOL; (* 印刷辊点动下降 *)
	i_xJogUp_Prn_G							: BOOL; (* 印刷辊点进上升  传动侧信号*)
	i_xJogDown_Prn_G						: BOOL; (* 印刷辊点动下降  传动侧信号*)
	i_xAllUp_Prn							: BOOL; (* 印刷辊整体上升 *)
	i_xAllDown_Prn							: BOOL; (* 印刷辊整体下降 *)
	i_xJogUp_Str_M							: BOOL; (* 张带辊点动上升 *)
	i_xJogDown_Str_M						: BOOL; (* 张带辊点动下降 *)
	i_xJogUp_Str_G							: BOOL; (* 张带辊点动上升  传动侧信号*)
	i_xJogDown_Str_G						: BOOL; (* 张带辊点动下降  传动侧信号*)
	i_xAllUp_Str							: BOOL; (* 张带辊整体上升 *)
	i_xAllDown_Str							: BOOL; (* 张带辊整体下降 *)
	i_xJogUp_Net_M							: BOOL; (* 网版辊点动前进 *)
	i_xJogDown_Net_M						: BOOL; (* 网版辊点动后退 *)
	i_xJogUp_Net_G							: BOOL; (* 网版辊点动前进 另传动侧信号*)
	i_xJogDown_Net_G						: BOOL; (* 网版辊点动后退  另传动侧信号*)
	i_xAllUp_Net							: BOOL; (* 网版辊整体前进 *)
	i_xAllDown_Net							: BOOL; (* 网版辊整体后退 *)

	i_xSuctionMotor							:BOOL; (* 吸风电机开关*)
	i_xNetMotor								:BOOL;(* 网辊电机开关*)
	i_xNetLock								:BOOL;(* 网辊锁紧开关*)
	i_xStop                             	:BOOL;(* 停止信号*)
	i_xRunning								:BOOL;(* 运行信号*)
	i_xNetPosLimit_Down						: BOOL; (* 网辊下限位 *)
	i_xPrnPosLimit_Up						: BOOL; (* 印刷辊上限位 *)
	i_xPrnPosLimit_Down						: BOOL; (* 印刷辊下限位 *)
	i_xPrnFastUp_M								: BOOL; (* 印刷辊快速上升 *)
	i_xPrnFastDown_M							: BOOL; (* 印刷辊快速下降 *)
	i_xHorzMotor_Alarm						: BOOL;(*横向报警*)
	(*新增变量-开始-wng.nt|2025.08.12.151630*)
	i_xPrnRollerLoose_H						: BOOL;(*夹板报警输入*)
	i_xLostPressure							: BOOL;(*气压低报警*)
	i_xPtcSignal							: BOOL;(*PTC过温报警*)

	i_xRsvd_DI0								: BOOL; (* 数字量输入保留0 *)
	i_xRsvd_DI1								: BOOL; (* 数字量输入保留1 *)
	i_xRsvd_DI2								: BOOL; (* 数字量输入保留2 *)
	i_xRsvd_DI3								: BOOL; (* 数字量输入保留3 *)
	i_xRsvd_DI4								: BOOL; (* 数字量输入保留4 *)
	i_xRsvd_DI5								: BOOL; (* 数字量输入保留5 *)
	i_xRsvd_DI6								: BOOL; (* 数字量输入保留6 *)
	i_xRsvd_DI7								: BOOL; (* 数字量输入保留7 *)
	i_xRsvd_DI8								: BOOL; (* 数字量输入保留8 *)
	i_xRsvd_DI9								: BOOL; (* 数字量输入保留9 *)
	i_wRsvd_AI0								: WORD; (* 模拟量输入保留0 *)
	i_wRsvd_AI1								: WORD; (* 模拟量输入保留1 *)
	i_wRsvd_AI2								: WORD; (* 模拟量输入保留2 *)
	i_wRsvd_AI3								: WORD; (* 模拟量输入保留3 *)
	i_wRsvd_AI4								: WORD; (* 模拟量输入保留4 *)
	i_wRsvd_AI5								: WORD; (* 模拟量输入保留5 *)

END_VAR
VAR_OUTPUT
	o_xEno									: BOOL;
	o_iErNo									: INT;

	o_xLamp_Linkage							: BOOL; (* 色组联动灯 *)
	o_xLamp_Inch							: BOOL; (* 单运行灯 *)
	o_xLamp_Estop							: BOOL; (* 急停灯输出 *)
	o_xLamp_Normal							: BOOL; (* 套色正常 *)
	o_xLamp_Warning							: BOOL; (* 套色报警 *)
	o_xLamp_Lost							: BOOL; (* 套色丢失 *)
	o_xLamp_AxisError						: BOOL; (* 轴故障指示 *)
	o_xRel_ArcAlarm_Unit					: BOOL; (* 本组套色报警输出 *)
	o_xLamp_Press							: BOOL; (* 合压指示 *)
	o_xRel_Press							: BOOL; (* 合压输出 *)
	o_xRel_UnPress							: BOOL; (* 离压输出 *)
	o_xHorzMotor_CW							: BOOL; (* 横向电机正转输出 *)
	o_xHorzMotor_CCW						: BOOL; (* 横向电机反转输出 *)
	o_xRel_Sleeve_Prn						: BOOL; (* 版辊套筒*)
	o_xRel_Sleeve_Net						: BOOL; (* 网辊套筒*)
	o_xRel_Plate_Push_Prn					: BOOL; (* 版辊推出*)
	o_xRel_Plate_Push_Net					: BOOL; (* 网辊推出*)
	o_xLamp_Inch_Net						: BOOL; (* 网辊单动灯 *)
	(*2024.09.28.094834//增加秦华IO*)
	o_xLamp_CorrctionPrn								: BOOL; (* 对版指示灯 *)
	o_xPM_Buzzer_Str								: BOOL; (* 张带辊装版蜂鸣器 *)
	o_xSuctionContactor								: BOOL; (* 吸风接触器 *)
	o_xDamMotorContactor								: BOOL; (* 润板电机接触器 *)
	o_xHydr_station_SV								: BOOL; (* 液压站电磁阀 *)

	//2026.05.21.161133
	o_xPrnRollerLoose_H						:BOOL;(*夹板松报警*)
	o_xLostPressure							:BOOL;(*气压低报警*)

	o_xRsvd_DO0								: BOOL; (* 数字量输出保留0 *)
	o_xRsvd_DO1								: BOOL; (* 数字量输出保留1 *)
	o_xRsvd_DO2								: BOOL; (* 数字量输出保留2 *)
	o_xRsvd_DO3								: BOOL; (* 数字量输出保留3 *)
	o_xRsvd_DO4								: BOOL; (* 数字量输出保留4 *)
	o_xRsvd_DO5								: BOOL; (* 数字量输出保留5 *)
	o_xRsvd_DO6								: BOOL; (* 数字量输出保留6 *)
	o_xRsvd_DO7								: BOOL; (* 数字量输出保留7 *)
	o_xRsvd_DO8								: BOOL; (* 数字量输出保留8 *)
	o_xRsvd_DO9								: BOOL; (* 数字量输出保留9 *)
	o_wRsvd_AO0								: WORD; (* 模拟量输出保留0 *)
	o_wRsvd_AO1								: WORD; (* 模拟量输出保留1 *)
	o_wRsvd_AO2								: WORD; (* 模拟量输出保留2 *)
	o_wRsvd_AO3								: WORD; (* 模拟量输出保留3 *)
	o_wRsvd_AO4								: WORD; (* 模拟量输出保留4 *)
	o_wRsvd_AO5								: WORD; (* 模拟量输出保留5 *)
END_VAR
VAR
END_VAR

{IMPLEMENTATION}
o_xEno:= i_xEn;
o_iErNo:= 0;
IF i_xEn THEN
	IF i_pstStIOMap_Axis_FE<>0 THEN
		IF i_xEnableInput THEN (* 输入 *)
			i_pstStIOMap_Axis_FE^.i_xLinkage					:= i_xLinkage; (* 联动 *)
			i_pstStIOMap_Axis_FE^.i_xInch					:= i_xInch; (* 单运行 *)
			i_pstStIOMap_Axis_FE^.i_xEstop					:= i_xEstop; (* 急停输入 *)
			i_pstStIOMap_Axis_FE^.i_xAlarmBell				:= i_xAlarmBell; (* 警报 *)
			i_pstStIOMap_Axis_FE^.i_xBigAdj					:= i_xBigAdj; (* 粗调 *)
			i_pstStIOMap_Axis_FE^.i_xLittleAdj				:= i_xLittleAdj; (* 细调 *)
			i_pstStIOMap_Axis_FE^.i_xPressMode_Auto			:= i_xPressMode_Auto; (* 自动合压 *)
			i_pstStIOMap_Axis_FE^.i_xPressMode_Manu			:= i_xPressMode_Manu; (* 手动合压 *)
			i_pstStIOMap_Axis_FE^.i_xPress					:= i_xPress; (* 合压输入 *)
			i_pstStIOMap_Axis_FE^.i_xUnPress					:= i_xUnPress; (* 离压输入 *)
			i_pstStIOMap_Axis_FE^.i_xUnPress_Inching			:= i_xUnPress_Inching; (* 点动离压 *)
			i_pstStIOMap_Axis_FE^.i_xMove_Up					:= i_xMove_Up; (* 上调 *)
			i_pstStIOMap_Axis_FE^.i_xMove_Down				:= i_xMove_Down; (* 下调 *)
			i_pstStIOMap_Axis_FE^.i_xMove_Left				:= i_xMove_Left; (* 左调 *)
			i_pstStIOMap_Axis_FE^.i_xMove_Right				:= i_xMove_Right; (* 右调 *)
			i_pstStIOMap_Axis_FE^.i_xPosLimit_Left			:= i_xPosLimit_Left; (* 左限位 *)
			i_pstStIOMap_Axis_FE^.i_xPosLimit_Right			:= i_xPosLimit_Right; (* 右限位 *)
			i_pstStIOMap_Axis_FE^.i_xHorzMotor_FastSpd		:= i_xHorzMotor_FastSpd; (* 横向电机快 *)
			i_pstStIOMap_Axis_FE^.i_xSleeve_Prn				:= i_xSleeve_Prn; (* 版辊套筒 *)
			i_pstStIOMap_Axis_FE^.i_xSleeve_Net				:= i_xSleeve_Net; (* 网辊套筒 *)
			i_pstStIOMap_Axis_FE^.i_xPlate_Push_Prn			:= i_xPlate_Push_Prn; (* 版辊推出 *)
			i_pstStIOMap_Axis_FE^.i_xPlate_Push_Net			:= i_xPlate_Push_Net; (* 网辊推出 *)

			i_pstStIOMap_Axis_FE^.i_xAcc						:= i_xAcc; (* 加速 *)
			i_pstStIOMap_Axis_FE^.i_xDec						:= i_xDec; (* 减速 *)
			i_pstStIOMap_Axis_FE^.i_xInch_Net				:= i_xInch_Net; (* 网棍云墨 *)
			(*2024.09.28.094834//增加秦华IO*)
			i_pstStIOMap_Axis_FE^.i_xJogPaper				:= i_xJogPaper; (* 走纸点动 *)
			i_pstStIOMap_Axis_FE^.i_xEn_Prn					:= i_xEn_Prn; (* 版辊使能开关 *)

			i_pstStIOMap_Axis_FE^.i_xPrnBigAdj				:= i_xPrnBigAdj; (* 印刷辊粗调 *)
			i_pstStIOMap_Axis_FE^.i_xPrnLittleAdj			:= i_xPrnLittleAdj; (* 印刷辊细调 *)
			i_pstStIOMap_Axis_FE^.i_xNetBigAdj				:= i_xNetBigAdj; (* 网辊粗调 *)
			i_pstStIOMap_Axis_FE^.i_xNetLittleAdj				:= i_xNetLittleAdj; (* 网辊细调 *)
			i_pstStIOMap_Axis_FE^.i_xStrBigAdj				:= i_xStrBigAdj; (* 张带辊粗调 *)
			i_pstStIOMap_Axis_FE^.i_xStrLittleAdj			:= i_xStrLittleAdj; (* 张带辊细调 *)

			i_pstStIOMap_Axis_FE^.i_xJogUp_Prn_M				:= i_xJogUp_Prn_M; (* 印刷辊点动上升 *)
			i_pstStIOMap_Axis_FE^.i_xJogDown_Prn_M			:= i_xJogDown_Prn_M; (* 印刷辊点动下降 *)
			i_pstStIOMap_Axis_FE^.i_xJogUp_Prn_G				:= i_xJogUp_Prn_G; (* 印刷辊点进上升 *)
			i_pstStIOMap_Axis_FE^.i_xJogDown_Prn_G			:= i_xJogDown_Prn_G; (* 印刷辊点动下降 *)
			i_pstStIOMap_Axis_FE^.i_xAllUp_Prn				:= i_xAllUp_Prn; (* 印刷辊整体上升 *)
			i_pstStIOMap_Axis_FE^.i_xAllDown_Prn				:= i_xAllDown_Prn; (* 印刷辊整体下降 *)
			i_pstStIOMap_Axis_FE^.i_xJogUp_Str_M				:= i_xJogUp_Str_M; (* 张带辊点动上升 *)
			i_pstStIOMap_Axis_FE^.i_xJogDown_Str_M			:= i_xJogDown_Str_M; (* 张带辊点动下降 *)
			i_pstStIOMap_Axis_FE^.i_xJogUp_Str_G				:= i_xJogUp_Str_G; (* 张带辊点动上升 *)
			i_pstStIOMap_Axis_FE^.i_xJogDown_Str_G			:= i_xJogDown_Str_G; (* 张带辊点动下降 *)
			i_pstStIOMap_Axis_FE^.i_xAllUp_Str				:= i_xAllUp_Str; (* 张带辊整体上升 *)
			i_pstStIOMap_Axis_FE^.i_xAllDown_Str				:= i_xAllDown_Str; (* 张带辊整体下降 *)
			i_pstStIOMap_Axis_FE^.i_xJogUp_Net_M				:= i_xJogUp_Net_M; (* 网版辊点动前进 *)
			i_pstStIOMap_Axis_FE^.i_xJogDown_Net_M			:= i_xJogDown_Net_M	; (* 网版辊点动后退 *)
			i_pstStIOMap_Axis_FE^.i_xJogUp_Net_G				:= i_xJogUp_Net_G; (* 网版辊点动前进 *)
			i_pstStIOMap_Axis_FE^.i_xJogDown_Net_G			:= i_xJogDown_Net_G; (* 网版辊点动后退 *)
			i_pstStIOMap_Axis_FE^.i_xAllUp_Net				:= i_xAllUp_Net; (* 网版辊整体前进 *)
			i_pstStIOMap_Axis_FE^.i_xAllDown_Net				:= i_xAllDown_Net; (* 网版辊整体后退 *)

			i_pstStIOMap_Axis_FE^.i_xSuctionMotor			:= i_xSuctionMotor; (* 吸风电机开关 *)
			i_pstStIOMap_Axis_FE^.i_xNetMotor				:= i_xNetMotor; (* 网辊电机开关 *)
			i_pstStIOMap_Axis_FE^.i_xNetLock					:= i_xNetLock; (* 网辊锁紧开关 *)
			i_pstStIOMap_Axis_FE^.i_xStop					:= i_xStop; (* 停止信号 *)
			i_pstStIOMap_Axis_FE^.i_xRunning					:= i_xRunning; (* 运行信号 *)
			i_pstStIOMap_Axis_FE^.i_xNetPosLimit_Down		:= i_xNetPosLimit_Down; (* 网辊下限位 *)
			i_pstStIOMap_Axis_FE^.i_xPrnPosLimit_Up			:= i_xPrnPosLimit_Up; (* 印刷辊上限位 *)
			i_pstStIOMap_Axis_FE^.i_xPrnPosLimit_Down		:= i_xPrnPosLimit_Down; (* 印刷辊下限位 *)
			i_pstStIOMap_Axis_FE^.i_xPrnFastUp_M				:= i_xPrnFastUp_M; (* 印刷辊快速上升 *)
			i_pstStIOMap_Axis_FE^.i_xPrnFastDown_M			:= i_xPrnFastDown_M; (* 印刷辊快速下降 *)
			i_pstStIOMap_Axis_FE^.i_xHorzMotor_Alarm			:=i_xHorzMotor_Alarm;
			(*新增变量-开始-wng.nt|2025.08.12.151630*)
			i_pstStIOMap_Axis_FE^.i_xPrnRollerLoose_H		:= i_xPrnRollerLoose_H;//				: BOOL;(*夹板报警输入*)
			i_pstStIOMap_Axis_FE^.i_xLostPressure	:= i_xLostPressure;//						: BOOL;(*气压低报警*)
			i_pstStIOMap_Axis_FE^.i_xPtcSignal		:= i_xPtcSignal;//				: BOOL;(*PTC过温报警*)

			i_pstStIOMap_Axis_FE^.i_xRsvd_DI0				:= i_xRsvd_DI0; (* 数字量输入保留0 *)
			i_pstStIOMap_Axis_FE^.i_xRsvd_DI1				:= i_xRsvd_DI1; (* 数字量输入保留1 *)
			i_pstStIOMap_Axis_FE^.i_xRsvd_DI2				:= i_xRsvd_DI2; (* 数字量输入保留2 *)
			i_pstStIOMap_Axis_FE^.i_xRsvd_DI3				:= i_xRsvd_DI3; (* 数字量输入保留3 *)
			i_pstStIOMap_Axis_FE^.i_xRsvd_DI4				:= i_xRsvd_DI4; (* 数字量输入保留4 *)
			i_pstStIOMap_Axis_FE^.i_xRsvd_DI5				:= i_xRsvd_DI5; (* 数字量输入保留5 *)
			i_pstStIOMap_Axis_FE^.i_xRsvd_DI6				:= i_xRsvd_DI6; (* 数字量输入保留6 *)
			i_pstStIOMap_Axis_FE^.i_xRsvd_DI7				:= i_xRsvd_DI7; (* 数字量输入保留7 *)
			i_pstStIOMap_Axis_FE^.i_xRsvd_DI8				:= i_xRsvd_DI8; (* 数字量输入保留8 *)
			i_pstStIOMap_Axis_FE^.i_xRsvd_DI9				:= i_xRsvd_DI9; (* 数字量输入保留9 *)
			i_pstStIOMap_Axis_FE^.i_wRsvd_AI0				:= i_wRsvd_AI0; (* 模拟量输入保留0 *)
			i_pstStIOMap_Axis_FE^.i_wRsvd_AI1				:= i_wRsvd_AI1; (* 模拟量输入保留1 *)
			i_pstStIOMap_Axis_FE^.i_wRsvd_AI2				:= i_wRsvd_AI2; (* 模拟量输入保留2 *)
			i_pstStIOMap_Axis_FE^.i_wRsvd_AI3				:= i_wRsvd_AI3; (* 模拟量输入保留3 *)
			i_pstStIOMap_Axis_FE^.i_wRsvd_AI4				:= i_wRsvd_AI4; (* 模拟量输入保留4 *)
			i_pstStIOMap_Axis_FE^.i_wRsvd_AI5				:= i_wRsvd_AI5; (* 模拟量输入保留5 *)

		END_IF

		IF i_xEnableOutput THEN (* 输出 *)
			o_xLamp_Linkage					:= i_pstStIOMap_Axis_FE^.o_xLamp_Linkage; (* 色组联动灯 *)
			o_xLamp_Inch					:= i_pstStIOMap_Axis_FE^.o_xLamp_Inch; (* 单运行灯 *)
			o_xLamp_Estop					:= i_pstStIOMap_Axis_FE^.o_xLamp_Estop; (* 急停灯输出 *)
			o_xLamp_Normal					:= i_pstStIOMap_Axis_FE^.o_xLamp_Normal; (* 套色正常 *)
			o_xLamp_Warning					:= i_pstStIOMap_Axis_FE^.o_xLamp_Warning; (* 套色报警 *)
			o_xLamp_Lost					:= i_pstStIOMap_Axis_FE^.o_xLamp_Lost; (* 套色丢失 *)
			o_xLamp_AxisError				:= i_pstStIOMap_Axis_FE^.o_xLamp_AxisError; (* 轴故障指示 *)
			o_xRel_ArcAlarm_Unit			:= i_pstStIOMap_Axis_FE^.o_xRel_ArcAlarm_Unit; (* 本组套色报警输出 *)
			o_xLamp_Press					:= i_pstStIOMap_Axis_FE^.o_xLamp_Press; (* 合压指示 *)
			o_xRel_Press					:= i_pstStIOMap_Axis_FE^.o_xRel_Press; (* 合压输出 *)
			o_xRel_UnPress					:= i_pstStIOMap_Axis_FE^.o_xRel_UnPress; (* 离压输出 *)
			o_xHorzMotor_CW					:= i_pstStIOMap_Axis_FE^.o_xHorzMotor_CW; (* 横向电机正转输出 *)
			o_xHorzMotor_CCW				:= i_pstStIOMap_Axis_FE^.o_xHorzMotor_CCW; (* 横向电机反转输出 *)
			o_xRel_Sleeve_Prn				:= i_pstStIOMap_Axis_FE^.o_xRel_Sleeve_Prn; (* 版辊套筒 *)
			o_xRel_Sleeve_Net				:= i_pstStIOMap_Axis_FE^.o_xRel_Sleeve_Net; (* 网辊套筒 *)
			o_xRel_Plate_Push_Prn			:= i_pstStIOMap_Axis_FE^.o_xRel_Plate_Push_Prn; (* 版辊推出 *)
			o_xRel_Plate_Push_Net			:= i_pstStIOMap_Axis_FE^.o_xRel_Plate_Push_Net; (* 网辊推出 *)
			o_xLamp_Inch_Net				:= i_pstStIOMap_Axis_FE^.o_xLamp_Inch_Net; (* 网辊云墨灯 *)
	(*2024.09.25.143257 增加io*)
			o_xLamp_CorrctionPrn			:= i_pstStIOMap_Axis_FE^.o_xLamp_CorrctionPrn; (* 对版指示灯 *)
			o_xPM_Buzzer_Str				:= i_pstStIOMap_Axis_FE^.o_xPM_Buzzer_Str; (* 张带辊装版蜂鸣器 *)
			o_xSuctionContactor				:= i_pstStIOMap_Axis_FE^.o_xSuctionContactor; (* 吸风接触器 *)
			o_xDamMotorContactor			:= i_pstStIOMap_Axis_FE^.o_xDamMotorContactor; (* 润板电机接触器 *)
			o_xHydr_station_SV				:= i_pstStIOMap_Axis_FE^.o_xHydr_station_SV; (* 液压站电磁阀 *)
	(*2026.05.21.161328*)
			o_xPrnRollerLoose_H				:=i_pstStIOMap_Axis_FE^.o_xPrnRollerLoose_H; (* 夹板松报警输出 *)
			o_xLostPressure					:=i_pstStIOMap_Axis_FE^.o_xLostPressure; (* 气压低报警输出 *)
	(*2026.01.26.155741//超旭用一下预留点位*)
			o_xRsvd_DO0						:= i_pstStIOMap_Axis_FE^.o_xRsvd_DO0; (* 数字量输出保留0 *)//充气电磁阀
			o_xRsvd_DO1						:= i_pstStIOMap_Axis_FE^.o_xRsvd_DO1; (* 数字量输出保留1 *)//墨盘电磁阀升
			o_xRsvd_DO2						:= i_pstStIOMap_Axis_FE^.o_xRsvd_DO2; (* 数字量输出保留2 *)//墨盘电磁阀降
			o_xRsvd_DO3						:= i_pstStIOMap_Axis_FE^.o_xRsvd_DO3; (* 数字量输出保留3 *)//墨盘锁轴电磁阀锁轴
			o_xRsvd_DO4						:= i_pstStIOMap_Axis_FE^.o_xRsvd_DO4; (* 数字量输出保留4 *)//墨盘锁轴电磁阀解锁
			o_xRsvd_DO5						:= i_pstStIOMap_Axis_FE^.o_xRsvd_DO5; (* 数字量输出保留5 *)//版辊电磁阀升锁轴
			o_xRsvd_DO6						:= i_pstStIOMap_Axis_FE^.o_xRsvd_DO6; (* 数字量输出保留6 *)//版辊电磁阀降解锁
			o_xRsvd_DO7						:= i_pstStIOMap_Axis_FE^.o_xRsvd_DO7; (* 数字量输出保留7 *)//停止灯（红）
			o_xRsvd_DO8						:= i_pstStIOMap_Axis_FE^.o_xRsvd_DO8; (* 数字量输出保留8 *)
			o_xRsvd_DO9						:= i_pstStIOMap_Axis_FE^.o_xRsvd_DO9; (* 数字量输出保留9 *)
			o_wRsvd_AO0						:= i_pstStIOMap_Axis_FE^.o_wRsvd_AO0; (* 模拟量输出保留0 *)
			o_wRsvd_AO1						:= i_pstStIOMap_Axis_FE^.o_wRsvd_AO1; (* 模拟量输出保留1 *)
			o_wRsvd_AO2						:= i_pstStIOMap_Axis_FE^.o_wRsvd_AO2; (* 模拟量输出保留2 *)
			o_wRsvd_AO3						:= i_pstStIOMap_Axis_FE^.o_wRsvd_AO3; (* 模拟量输出保留3 *)
			o_wRsvd_AO4						:= i_pstStIOMap_Axis_FE^.o_wRsvd_AO4; (* 模拟量输出保留4 *)
			o_wRsvd_AO5						:= i_pstStIOMap_Axis_FE^.o_wRsvd_AO5; (* 模拟量输出保留5 *)
		END_IF
	ELSE
		o_iErNo:= -1;
	END_IF
ELSE
	o_xLamp_Linkage					:= FALSE; (* 色组联动灯 *)
	o_xLamp_Inch					:= FALSE; (* 单运行灯 *)
	o_xLamp_Estop					:= FALSE; (* 急停灯输出 *)
	o_xLamp_Normal					:= FALSE; (* 套色正常 *)
	o_xLamp_Warning					:= FALSE; (* 套色报警 *)
	o_xLamp_Lost					:= FALSE; (* 套色丢失 *)
	o_xLamp_AxisError				:= FALSE; (* 轴故障指示 *)
	o_xRel_ArcAlarm_Unit			:= FALSE; (* 本组套色报警输出 *)
	o_xLamp_Press					:= FALSE; (* 合压指示 *)
	o_xRel_Press					:= FALSE; (* 合压输出 *)
	o_xRel_UnPress					:= FALSE; (* 离压输出 *)
	o_xHorzMotor_CW					:= FALSE; (* 横向电机正转输出 *)
	o_xHorzMotor_CCW				:= FALSE; (* 横向电机反转输出 *)
	o_xRel_Sleeve_Prn				:= FALSE; (* 版辊套筒 *)
	o_xRel_Sleeve_Net				:= FALSE; (* 网辊套筒 *)
	o_xRel_Plate_Push_Prn			:= FALSE; (* 版辊推出 *)
	o_xRel_Plate_Push_Net			:= FALSE; (* 网辊推出 *)

	o_xRsvd_DO0						:= FALSE; (* 数字量输出保留0 *)
	o_xRsvd_DO1						:= FALSE; (* 数字量输出保留1 *)
	o_xRsvd_DO2						:= FALSE; (* 数字量输出保留2 *)
	o_xRsvd_DO3						:= FALSE; (* 数字量输出保留3 *)
	o_xRsvd_DO4						:= FALSE; (* 数字量输出保留4 *)
	o_xRsvd_DO5						:= FALSE; (* 数字量输出保留5 *)
	o_xRsvd_DO6						:= FALSE; (* 数字量输出保留6 *)
	o_xRsvd_DO7						:= FALSE; (* 数字量输出保留7 *)
	o_xRsvd_DO8						:= FALSE; (* 数字量输出保留8 *)
	o_xRsvd_DO9						:= FALSE; (* 数字量输出保留9 *)
	o_wRsvd_AO0						:= 0; (* 模拟量输出保留0 *)
	o_wRsvd_AO1						:= 0; (* 模拟量输出保留1 *)
	o_wRsvd_AO2						:= 0; (* 模拟量输出保留2 *)
	o_wRsvd_AO3						:= 0; (* 模拟量输出保留3 *)
	o_wRsvd_AO4						:= 0; (* 模拟量输出保留4 *)
	o_wRsvd_AO5						:= 0; (* 模拟量输出保留5 *)
END_IF
